(* IEC 61131-3 sources: daoli-st-library/DL_Device (part 20) *)

(* ---- FB_DL_EfEmDoorInterlockPlus.st ---- *)
(*==============================================================================
 * 组件名称 (Component)  : FB_DL_EfEmDoorInterlockPlus
 * 所属子库 (Sublibrary) : DL_Device
 * 当前版本 (Version)    : 1.0.0
 * 兼容性 (Platform)     : CODESYS 3.5 / TwinCAT 3 / 汇川 InoProShop（纯标准元素，零方言）
 * 功能描述 (Function)   : EFEM 门 / 阀 / 真空三域互斥与首因仲裁。唯一放行出口 bRelease
 *                         由四类阻断条件（门未关、阀位矛盾、真空不足、片在位）合成，阻断
 *                         域掩码逐域可见，首因只报一个编号（同拍取编号最小，锁存至复位）。
 *                         不做门体驱动输出、不做真空泵控制、不做安全回路硬线替代（安全
 *                         回路必须另有硬线双通道，本件只做逻辑侧互斥）。
 *                         门状态字位段（头注释即契约）：bit0 门关到位 ｜ bit1 门开到位 ｜
 *                         bit2 门锁到位 ｜ bit3~bit15 保留且必须为 0。
 * 溯源 (Origin)         : 道莅 clean-room 防御性实现
 * 本文件内含 (Contains) : TYPE E_DL_EfEmDomain / FUNCTION_BLOCK FB_DL_EfEmDoorInterlockPlus
 * 依赖 (Depends)        : 无（纯布尔/浮点防御逻辑，仅 Standard.library 的 ABS）
 * 红线自检 (Redline)    : 无外部全局变量、无硬件地址直引 ｜ 全变量中英双语同行注释
 *                         真空门限判零防除零 ｜ 真空非有限按保守侧（真空不足）处理 ｜
 *                         阀位矛盾判定前置于互斥仲裁 ｜ 枚举显式赋值 ｜ CASE 含 ELSE 兜底
 *                         本件无定时器/沿实例，故无周期刷新项（结构上无条件分支）
 * 错误码表 (Codes)      : 16#0003_03AC 就绪（放行或禁用，无故障）
 *                         16#0003_03AD 故障级 门状态字非法（保留位非 0）。反证句：保留位
 *                                    脏数据在输出侧与「门未关」同为禁行，不可由首因 1 区分，
 *                                    故必须独立成码
 *                         16#0003_03AE 故障级 阀位矛盾或真空门限组态非法（双反馈同 TRUE /
 *                                    同为 FALSE / 门限 ≤0）
 *                         16#0003_03AF 故障级 真空读数非有限，按「真空不足」保守侧禁行
 *                         16#0003_03B0 预留：本版不发码（下一轮区间起点，禁止回填）
 * 修订历史 (Revision)   : 2026-11-17  v1.0.0  首版入库 · R28 · 阶段三批 1
 * 验收向量 (Acceptance) : 正向 门关（状态字 bit0=1、bit2=1）、阀开反馈有效、真空 0.1 kPa
 *                         低于门限 5 kPa → 禁行、首因 3、掩码 bit2；抽到 0.05 kPa →
 *                         放行、首因清零
 *                         反向 阀双反馈同为 FALSE → 16#0003_03AE 且禁行；真空给 NaN →
 *                         16#0003_03AF 且按真空不足禁行（首因 3）；门限给 0 → 16#0003_03AE；
 *                         状态字保留位 bit7 置 1 → 16#0003_03AD 且禁行
 *============================================================================*)

(*-----------------------------------------------------------------------------
 * 枚举: E_DL_EfEmDomain（归属本功能块，同文件发布，全库唯一定义）
 * 含义: 首因所属域，每个成员在 CASE 中有且仅有一个标签。
 *----------------------------------------------------------------------------*)
TYPE E_DL_EfEmDomain :
(
    eNone    := 0,    // 无阻断域：三域全放行 / No blocking domain, all domains released
    eDoor    := 1,    // 门域：门未关到位 / Door domain, the door is not closed
    eValve   := 2,    // 阀域：阀位矛盾 / Valve domain, contradictory valve position
    eVacuum  := 3,    // 真空域：真空不足或读数非有限 / Vacuum domain, insufficient vacuum or a non-finite reading
    eWafer   := 4,    // 片域：腔内片在位（E84 语义） / Wafer domain, a wafer is present inside the chamber
    eIllegal := 99    // 非法域：状态字保留位非 0 / Illegal domain, reserved bits of the status word are set
);
END_TYPE

FUNCTION_BLOCK FB_DL_EfEmDoorInterlockPlus
VAR_INPUT
    bEnable         : BOOL := FALSE;      // 使能，FALSE 即禁行（失效导向安全侧） / Enable, FALSE forces the release output off
    uDoorStatusWord : WORD;               // 门状态字 [bit]，bit0 关到位 bit1 开到位 bit2 锁到位 bit3~15 保留 / Door status word
    bValveClosed    : BOOL := FALSE;      // 阀关到位反馈 / Valve closed feedback
    bValveOpened    : BOOL := FALSE;      // 阀开到位反馈 / Valve opened feedback
    fVacuum_kPa     : REAL := 101.3;      // 腔体真空 [kPa(abs)]，域 0~101.3 / Chamber vacuum in kilopascal absolute, domain 0 to 101.3
    fVacuumOk_kPa   : REAL := 5.0;        // 允许开门真空门限 [kPa(abs)] / Vacuum threshold permitting the door to open
    bWaferPresent   : BOOL := FALSE;      // 腔内片在位（E84 语义） / Wafer present in the chamber
    bReset          : BOOL := FALSE;      // 首因与锁存复位，上升沿生效 / First-cause and latch reset, rising edge
END_VAR
VAR_OUTPUT
    bRelease        : BOOL;               // 三域放行（唯一出口） / Three-domain release, the single outlet
    bDoorPermit     : BOOL;               // 允许开门（与放行同源，语义收窄为门域） / Door open permit, same source as the release
    uFirstCause     : UINT;               // 首因编号 1 门未关 2 阀位矛盾 3 真空不足 4 片在位 [—] / First cause number
    uBlockMask      : WORD;               // 阻断域掩码 bit0 门 bit1 阀 bit2 真空 bit3 片 [bit] / Blocking domain mask
    bError          : BOOL;               // 故障级标志，仅故障级码置位 / Fault-class flag, set on fault codes only
    eErr            : UDINT;              // 错误码，段位 16#0003_xxxx / Error code in segment 16#0003_xxxx
END_VAR
VAR
    _bInit          : BOOL := FALSE;      // 首扫标志，取非判定 / First-scan flag, tested negated
    _bDoorClosed    : BOOL;               // 门关到位（状态字 bit0） / Door closed, status word bit 0
    _bLocked        : BOOL;               // 门锁到位（状态字 bit2） / Door locked, status word bit 2
    _bReservedBad   : BOOL;               // 状态字保留位非 0 / Reserved bits of the status word are set
    _bValveBad      : BOOL;               // 阀位矛盾 / Contradictory valve position
    _bVacBad        : BOOL;               // 真空不足（含读数非有限） / Insufficient vacuum including non-finite readings
    _bCfgBad        : BOOL;               // 真空门限组态非法 / Vacuum threshold configuration invalid
    _bBlkDoor       : BOOL;               // 门域阻断 / Door domain blocked
    _bBlkValve      : BOOL;               // 阀域阻断 / Valve domain blocked
    _bBlkVac        : BOOL;               // 真空域阻断 / Vacuum domain blocked
    _bBlkWafer      : BOOL;               // 片域阻断 / Wafer domain blocked
    _bAnyBlock      : BOOL;               // 任一域阻断 / Any domain blocked
    _bFirstLatched  : BOOL;               // 首因已锁存（锁存后不再改判） / First cause latched and no longer re-arbitrated
    _eDomain        : E_DL_EfEmDomain := E_DL_EfEmDomain.eNone; // 当前首因域 / Current first-cause domain
    _rtrigReset     : R_TRIG;             // 复位上升沿 / Rising edge of the reset command
END_VAR
VAR CONSTANT
    DL_EFEM_READY      : UDINT := 16#0003_03AC;  // 就绪码 / Ready code
    DL_EFEM_WORD_BAD   : UDINT := 16#0003_03AD;  // 故障级状态字非法码 / Fault code for an illegal status word
    DL_EFEM_VALVE_BAD  : UDINT := 16#0003_03AE;  // 故障级阀位矛盾或组态非法码 / Fault code for a valve contradiction or bad configuration
    DL_EFEM_VAC_BAD    : UDINT := 16#0003_03AF;  // 故障级真空非有限码 / Fault code for a non-finite vacuum reading
    DL_EFEM_VAC_LO     : REAL := 0.0;            // 真空物理下限 [kPa(abs)] / Physical vacuum lower bound
    DL_EFEM_VAC_HI     : REAL := 101.3;          // 真空物理上限 [kPa(abs)] / Physical vacuum upper bound
    DL_EFEM_MASK_DOOR  : WORD := 16#0001;        // 门域掩码位 [bit] / Door domain mask bit
    DL_EFEM_MASK_VALVE : WORD := 16#0002;        // 阀域掩码位 [bit] / Valve domain mask bit
    DL_EFEM_MASK_VAC   : WORD := 16#0004;        // 真空域掩码位 [bit] / Vacuum domain mask bit
    DL_EFEM_MASK_WAFER : WORD := 16#0008;        // 片域掩码位 [bit] / Wafer domain mask bit
    DL_EFEM_WORD_RSV   : WORD := 16#FFF8;        // 状态字保留位掩码 [bit] / Reserved bit mask of the status word
    DL_EFEM_CAUSE_DOOR : UINT := 1;               // 首因 1 门未关 / First cause 1, the door is not closed
    DL_EFEM_CAUSE_VALVE : UINT := 2;              // 首因 2 阀位矛盾 / First cause 2, contradictory valve position
    DL_EFEM_CAUSE_VAC  : UINT := 3;               // 首因 3 真空不足 / First cause 3, insufficient vacuum
    DL_EFEM_CAUSE_WAFER : UINT := 4;              // 首因 4 片在位 / First cause 4, a wafer is present
END_VAR

// 段 1｜输出与单拍标志预置（放行类输出先清零：失效导向安全侧）
bRelease := FALSE;                                  // 放行出口先清 / Release outlet cleared first
bDoorPermit := FALSE;                               // 开门许可先清 / Door permit cleared first
uFirstCause := 0;                                   // 首因预清 / First cause pre-cleared
uBlockMask := 16#0000;                              // 掩码预清 / Mask pre-cleared
bError := FALSE;                                    // 故障标志预清 / Fault flag pre-cleared
eErr := 0;                                          // 错误码预清 / Error code pre-cleared

// 段 2｜沿检测无条件周期刷新（严禁置于分支内）
_rtrigReset(CLK := bReset);                         // 复位沿 / Reset edge

// 段 3｜首扫初始化（判据取非，R19）
IF NOT _bInit THEN
    _eDomain := E_DL_EfEmDomain.eNone;              // 首因域待机 / First-cause domain starts at none
    _bInit := TRUE;                                 // 首扫只做一次 / The first scan runs once
END_IF

// 段 4｜复位路径：清首因锁存（放行条件本身不清，条件仍在则同拍重新锁存）
IF _rtrigReset.Q THEN
    _bFirstLatched := FALSE;                        // 首因锁存解除 / First-cause latch released
    uFirstCause := 0;                               // 首因编号清 / First-cause number cleared
    _eDomain := E_DL_EfEmDomain.eNone;              // 首因域清 / First-cause domain cleared
END_IF

// 段 5｜门状态字解析（保留位脏数据先判，避免位段错位被当门未关）
_bDoorClosed := (uDoorStatusWord AND DL_EFEM_MASK_DOOR) <> 16#0000;   // bit0 关到位 / Bit 0, closed position reached
_bLocked := (uDoorStatusWord AND 16#0004) <> 16#0000;                 // bit2 锁到位 / Bit 2, locking position reached
_bReservedBad := (uDoorStatusWord AND DL_EFEM_WORD_RSV) <> 16#0000;   // 保留位非 0 / Reserved bits are set

// 段 6｜阀位矛盾闸（前置于互斥仲裁：矛盾状态下首因必须指阀域而不是门域）
_bValveBad := (bValveClosed AND bValveOpened) OR ((NOT bValveClosed) AND (NOT bValveOpened));

// 段 7｜真空组态与读数闸（门限判零防除零；读数非有限按真空不足保守侧）
_bCfgBad := (fVacuumOk_kPa <> fVacuumOk_kPa) OR ((fVacuumOk_kPa - fVacuumOk_kPa) <> (fVacuumOk_kPa - fVacuumOk_kPa))
         OR (fVacuumOk_kPa <= DL_EFEM_VAC_LO) OR (fVacuumOk_kPa > DL_EFEM_VAC_HI);
IF (fVacuum_kPa <> fVacuum_kPa) OR ((fVacuum_kPa - fVacuum_kPa) <> (fVacuum_kPa - fVacuum_kPa)) THEN
    _bVacBad := TRUE;                               // 读数非有限：按真空不足处理 / Non-finite reading treated as insufficient vacuum
    eErr := DL_EFEM_VAC_BAD;                        // 故障级：真空读数非有限 / Fault, non-finite vacuum reading
    bError := TRUE;
ELSE
    _bVacBad := (fVacuum_kPa > fVacuumOk_kPa);      // 真空值高于门限 = 真空不足 / A value above the threshold means insufficient vacuum
END_IF
IF _bCfgBad THEN
    eErr := DL_EFEM_VALVE_BAD;                      // 故障级：真空门限组态非法 / Fault, the vacuum threshold configuration is invalid
    bError := TRUE;
END_IF
IF _bReservedBad THEN
    eErr := DL_EFEM_WORD_BAD;                       // 故障级：状态字保留位非 0 / Fault, reserved bits of the status word are set
    bError := TRUE;
END_IF
IF _bValveBad THEN
    eErr := DL_EFEM_VALVE_BAD;                      // 故障级：阀位矛盾（先于互斥判定） / Fault, contradictory valve position checked before the arbitration
    bError := TRUE;
END_IF

// 段 8｜四域阻断判定（掩码逐域可见，首因只报一个）
_bBlkDoor := (NOT _bDoorClosed) OR (NOT _bLocked);  // 门域：关到位与锁到位缺一即阻断 / Door domain blocked unless closed and locked
_bBlkValve := _bValveBad OR _bCfgBad;               // 阀域：阀位矛盾或组态非法即阻断 / Valve domain blocked on a contradiction or bad configuration
_bBlkVac := _bVacBad OR _bCfgBad;                   // 真空域：真空不足或组态非法即阻断 / Vacuum domain blocked on insufficient vacuum or bad configuration
_bBlkWafer := bWaferPresent;                        // 片域：腔内片在位即阻断 / Wafer domain blocked while a wafer is present
_bAnyBlock := _bBlkDoor OR _bBlkValve OR _bBlkVac OR _bBlkWafer;   // 任一域阻断 / Any domain blocked
IF _bBlkDoor THEN
    uBlockMask := uBlockMask OR DL_EFEM_MASK_DOOR;  // 门域掩码置位 / Door domain mask bit set
END_IF
IF _bBlkValve THEN
    uBlockMask := uBlockMask OR DL_EFEM_MASK_VALVE; // 阀域掩码置位 / Valve domain mask bit set
END_IF
IF _bBlkVac THEN
    uBlockMask := uBlockMask OR DL_EFEM_MASK_VAC;   // 真空域掩码置位 / Vacuum domain mask bit set
END_IF
IF _bBlkWafer THEN
    uBlockMask := uBlockMask OR DL_EFEM_MASK_WAFER; // 片域掩码置位 / Wafer domain mask bit set
END_IF

// 段 9｜首因仲裁（仅未锁存时仲裁；顺序 1→4 即同拍取编号最小）
IF (NOT _bFirstLatched) AND _bAnyBlock THEN
    IF _bBlkDoor THEN
        _eDomain := E_DL_EfEmDomain.eDoor;          // 优先 1：门未关 / Priority 1, the door is not closed
    ELSIF _bBlkValve THEN
        _eDomain := E_DL_EfEmDomain.eValve;         // 优先 2：阀位矛盾 / Priority 2, contradictory valve position
    ELSIF _bBlkVac THEN
        _eDomain := E_DL_EfEmDomain.eVacuum;        // 优先 3：真空不足 / Priority 3, insufficient vacuum
    ELSE
        _eDomain := E_DL_EfEmDomain.eWafer;         // 优先 4：片在位 / Priority 4, a wafer is present
    END_IF
    _bFirstLatched := TRUE;                         // 首因锁存 / First cause latched
ELSIF (NOT _bAnyBlock) THEN
    _bFirstLatched := FALSE;                        // 阻断全消失：锁存解除（状态量随条件销号） / All blocks cleared, the latch is released
    _eDomain := E_DL_EfEmDomain.eNone;              // 首因域回无 / First-cause domain back to none
END_IF

// 段 10｜首因域映射（ENUM + CASE + ELSE 兜底）
CASE _eDomain OF
    E_DL_EfEmDomain.eNone:
        uFirstCause := 0;                           // 无首因 / No first cause
    E_DL_EfEmDomain.eDoor:
        uFirstCause := DL_EFEM_CAUSE_DOOR;          // 首因 1 / First cause 1
    E_DL_EfEmDomain.eValve:
        uFirstCause := DL_EFEM_CAUSE_VALVE;         // 首因 2 / First cause 2
    E_DL_EfEmDomain.eVacuum:
        uFirstCause := DL_EFEM_CAUSE_VAC;           // 首因 3 / First cause 3
    E_DL_EfEmDomain.eWafer:
        uFirstCause := DL_EFEM_CAUSE_WAFER;         // 首因 4 / First cause 4
    E_DL_EfEmDomain.eIllegal:
        uFirstCause := 0;                           // 非法域不报首因，由 03AD 表达 / The illegal domain reports no first cause, 03AD carries it
        eErr := DL_EFEM_WORD_BAD;                   // 故障级：非法域 / Fault, illegal domain
        bError := TRUE;
    ELSE
        // 非法枚举值兜底（故障级，状态字非法码承载）
        uFirstCause := 0;
        eErr := DL_EFEM_WORD_BAD;                   // 故障级：枚举越界 / Fault, the enumeration is out of range
        bError := TRUE;
        _eDomain := E_DL_EfEmDomain.eIllegal;
END_CASE

// 段 11｜放行出口（唯一出口；使能跌落即禁行，故障级存在亦禁行）
bRelease := bEnable AND (NOT _bAnyBlock) AND (NOT _bReservedBad) AND (NOT _bCfgBad) AND (NOT _bValveBad) AND (NOT _bVacBad);
bDoorPermit := bRelease;                            // 开门许可与放行同源 / Door permit shares the release source
IF bRelease THEN
    eErr := DL_EFEM_READY;                          // 就绪：三域放行 / Ready, all domains released
ELSE
    IF NOT bEnable THEN
        eErr := DL_EFEM_READY;                      // 禁用为正常停机（掩码已标全阻断域） / Disable is a normal stop, the mask shows the blocked domains
    END_IF
END_IF
END_FUNCTION_BLOCK

(* ---- FB_DL_ElectricLinearActuator.st ---- *)
(*
  ==================================================================
  组件名 Component  : FB_DL_ElectricLinearActuator
  分类   Category   : DL_Device
  复杂度 Complexity  : cx5
  版本   Version    : 1.0.0
  功能   Purpose    : 电动推杆驱动。无位置反馈，纯时间 / 电流双模到位判定：
                      限位开关反馈模（任一端限位反馈触发）与电流堵转模（电
                      流持续超堵转阈值 tStallDebounce 消抖判到位）并联，任
                      一判据先到即停并锁存到位指示；硬过流立即脱扣；全程
                      超时保护；双输出互锁绝不同得电。
  来源   Source     : t2-2-lbp（三段分层骨架）
  溯源   Origin     : IEC 61131-3 标准语义的道莅防御性实现；电动推杆堵转
                      电流判到位与限位互锁为行业公知工程语义，clean-room
                      自研实现，未复制 LBP 或任何厂商私有库源码。
  平台   Platform   : 纯 IEC 61131-3（Standard.library: TON / R_TRIG，无私有库）
  分工声明 Split     : 与 DL_Device 存量 FB_DL_DolMotor / FB_DL_SoftStarterDrive
                      分工——两者为电机启动家族（驱动器封装），本件为直线
                      执行机构（推杆本体行程与堵转管理），不做接触器 / 晶闸
                      管启动家族语义。
  作者   Author     : 道莅代码库 · PLC 编程专家（R58）
  ------------------------------------------------------------------
  边界 Boundary     :
                      一 组态域：fCurNomA > 0（非有限闸覆盖），fCurStallMul
                         > 1.0，fCurHiMul > fCurStallMul（硬过流阈值高于堵转
                         阈值，R100 配比约束），tStrokeMax > T#0S，tStallDebounce
                         ≥ T#0S（取零为电流模禁用，仅限位模）；
                      二 双模并联：限位反馈与电流堵转任一先到即到位停机，
                         到位指示锁存至反向运动或复位沿；
                      三 双命令同拍拒绝（复位优先 = 安全侧不动作，静默拒
                         绝不置故障，本拍双输出全断）；
                      四 运动相电流非有限（R151 组态域闸全覆盖）判传感失效
                         故障级；复位沿作用域：清故障锁存 / 清到位指示 / 迁
                         空闲（三项逐项声明，解除路径 = bReset 上升沿 R188）；
                      五 无全局变量、无外部变量声明、无物理地址寻址。
  修订记录 Revision  :
    2026-11-21  v1.0.0  R58 首版（批 2 · 序号 8）
  ==================================================================
*)

TYPE E_DL_ElaPhase :
(
    eElaIdle := 0,  // 空闲：消化命令，双输出断开 / idle, both outputs off
    eElaExt  := 10, // 伸出中：正转输出得电 / extending, the forward output on
    eElaRet  := 20, // 缩回中：反转输出得电 / retracting, the reverse output on
    eElaFault:= 90  // 故障锁存：双输出安全侧断开 / the latched fault, both outputs off on the safe side
);
END_TYPE

TYPE E_DL_ElaCause :
(
    eNone          := 0, // 无成因 / no cause
    eCfgBad        := 1, // 组态非法：电流标称 / 倍数配比 / 时间窗越域（故障级，与 bError 配对）/ an illegal config
    eCurBad        := 2, // 运动相电流非有限（传感失效，故障级，与 bError 配对）/ a non finite current in motion
    eCurOverHard   := 3, // 硬过流立即脱扣（故障级，与 bError 配对）/ a hard overcurrent trip
    eStrokeTimeout := 4, // 全程超时（故障级，与 bError 配对）/ a stroke timeout
    ePhaseBad      := 5  // 非法相位兜底（故障级，与 bError 配对）/ an illegal phase fallback
);
END_TYPE

FUNCTION_BLOCK FB_DL_ElectricLinearActuator
VAR_INPUT
    bCmdExt        : BOOL := FALSE;  // 伸出命令电平 [-] / the extend command level
    bCmdRet        : BOOL := FALSE;  // 缩回命令电平 [-] / the retract command level
    bLimExtFbk     : BOOL := FALSE;  // 伸出限位开关反馈，TRUE = 已达伸出端 [-] / the extend limit feedback, true = at the extend end
    bLimRetFbk     : BOOL := FALSE;  // 缩回限位开关反馈，TRUE = 已达缩回端 [-] / the retract limit feedback, true = at the retract end
    fMotCurA       : LREAL := 0.0;   // 电机电流实测 [安培] / the motor current actual [ampere]
    fCurNomA       : LREAL := 4.0;   // 标称运行电流 [安培]，域 大于 0 / the nominal running current [ampere], above zero
    fCurStallMul   : LREAL := 1.5;   // 堵转判定倍数 [倍]，域 大于 1.0 / the stall verdict multiplier, above one
    fCurHiMul      : LREAL := 2.5;   // 硬过流倍数 [倍]，域 大于堵转倍数 / the hard overcurrent multiplier, above the stall multiplier
    tStrokeMax     : TIME := T#30S;  // 全程最大时间窗 [毫秒] / the full stroke max window [millisecond]
    tStallDebounce : TIME := T#300MS; // 堵转消抖窗 [毫秒]，取零禁用电流模 / the stall debounce window, zero disables the current mode
    bEnable        : BOOL := TRUE;   // 使能，失能双输出安全侧断开并迁空闲 [-] / enable, disabling opens both outputs and returns idle
    bReset         : BOOL := FALSE;  // 复位上升沿清故障锁存 [-] / reset rising edge clears the fault latch
END_VAR
VAR_OUTPUT
    bOutExt   : BOOL := FALSE; // 电机正转输出（仅伸出相）[-] / the forward output, the extend phase only
    bOutRet   : BOOL := FALSE; // 电机反转输出（仅缩回相）[-] / the reverse output, the retract phase only
    bInPosExt : BOOL := FALSE; // 伸出到位指示（锁存至反向或复位）[-] / the extend in position latch
    bInPosRet : BOOL := FALSE; // 缩回到位指示（锁存至反向或复位）[-] / the retract in position latch
    bArrByCur : BOOL := FALSE; // 本次到位由电流堵转模判定的指示 [-] / the arrival by the current mode indicator
    ePhase    : E_DL_ElaPhase := E_DL_ElaPhase.eElaIdle; // 相位出口 [枚举] / the phase outlet
    eCause    : E_DL_ElaCause := E_DL_ElaCause.eNone; // 成因出口，锁存回放 [枚举] / the cause outlet replayed
    bError    : BOOL := FALSE; // 故障锁存标志 [-] / the fault latch flag
END_VAR
VAR
    rtReset  : R_TRIG; // 复位沿检测，段 0 无条件刷新 / the reset edge
    tonStroke: TON;    // 全程时间窗，段 0 无条件刷新 / the stroke window
    tonStall : TON;    // 堵转消抖窗，段 0 无条件刷新 / the stall debounce window
    _ePhase  : E_DL_ElaPhase := E_DL_ElaPhase.eElaIdle; // 内部相位，CASE 唯一写入目标 / the internal phase
    _eFaulC  : E_DL_ElaCause := E_DL_ElaCause.eNone; // 故障级成因，锁存至复位沿 / the fault cause latched
    _bFault  : BOOL := FALSE; // 故障锁存位 [-] / the fault latch bit
    _bCfgOk  : BOOL := FALSE; // 组态域内 [-] / the config inside the domain
    _bInit   : BOOL := FALSE; // 首扫初始化完成标志（R310）/ the first scan flag
    _lrStall : LREAL;  // 堵转电流阈值工作量 [安培] / the stall threshold work value
    _lrHi    : LREAL;  // 硬过流阈值工作量 [安培] / the hard overcurrent threshold work value
END_VAR

// 段 0｜定时器与沿检测无条件周期刷新（禁入分支，FB50-1）/ segment 0, the unconditional refresh
rtReset(CLK := bReset); // 复位沿 / the reset edge
tonStroke(IN := ((_ePhase = E_DL_ElaPhase.eElaExt) OR (_ePhase = E_DL_ElaPhase.eElaRet)) AND (NOT _bFault) AND bEnable, PT := tStrokeMax); // 全程窗，IN 串载能相闸（纯相驻留，R145）/ the stroke window on the powered phases
tonStall(IN := ((_ePhase = E_DL_ElaPhase.eElaExt) OR (_ePhase = E_DL_ElaPhase.eElaRet)) AND (NOT _bFault) AND bEnable AND (_lrStall > 0.0) AND (fMotCurA > _lrStall), PT := tStallDebounce); // 堵转消抖窗（电流模使能且超阈）/ the stall debounce window, the current mode enabled and above the threshold

// 段 1｜首扫初始化（R310）/ segment 1, the first scan
IF NOT _bInit THEN // 首扫一拍 / the first scan
    _bInit := TRUE; // 置首扫标志 / raise the flag
END_IF

// 段 2｜复位沿作用域：清故障锁存 / 清到位指示 / 迁空闲（三项逐项声明，边界四）/ segment 2, the reset edge scope
IF rtReset.Q THEN // 复位沿 / the reset edge
    _bFault := FALSE; // 作用域一：清故障锁存 / scope one, clear the fault latch
    _eFaulC := E_DL_ElaCause.eNone; // 作用域一：清成因 / scope one, clear the cause
    bInPosExt := FALSE; // 作用域二：清伸出到位 / scope two, clear the extend latch
    bInPosRet := FALSE; // 作用域二：清缩回到位 / scope two, clear the retract latch
    bArrByCur := FALSE; // 作用域二：清电流模指示 / scope two, clear the current mode flag
    _ePhase := E_DL_ElaPhase.eElaIdle; // 作用域三：迁空闲相 / scope three, back to idle
END_IF

// 段 3｜组态域闸（边界一，R151 全覆盖：电流标称非有限 + 倍数配比 + 时间窗）/ segment 3, the config gate
_bCfgOk := (fCurNomA = fCurNomA) AND ((fCurNomA - fCurNomA) = (fCurNomA - fCurNomA)) // 标称电流非有限双判据 / the nominal current finiteness
        AND (fCurNomA > 0.0) // 标称电流域 / the nominal domain
        AND (fCurStallMul > 1.0) // 堵转倍数域 / the stall multiplier domain
        AND (fCurHiMul > fCurStallMul) // 硬过流高于堵转配比（R100）/ the hard above the stall pairing
        AND (tStrokeMax > T#0S) // 全程窗域 / the stroke window domain
        AND (tStallDebounce >= T#0S); // 消抖窗域（零 = 电流模禁用）/ the debounce domain, zero disables the current mode
IF NOT _bCfgOk THEN // 组态越域 / a config violation
    IF NOT _bFault THEN // 未锁存才迁移（锁存回放 R152）/ migrate only while unlatched
        _bFault := TRUE; // 置故障锁存 / raise the fault latch
        _eFaulC := E_DL_ElaCause.eCfgBad; // 故障级成因（R45 配对）/ the fault cause
        _ePhase := E_DL_ElaPhase.eElaFault; // 迁故障相（锁存与迁相同分支，FB50-1）/ migrate to the fault phase
    END_IF
END_IF
_lrStall := fCurNomA * fCurStallMul; // 堵转阈值（组态闸已证有限正值）/ the stall threshold
_lrHi := fCurNomA * fCurHiMul; // 硬过流阈值 / the hard threshold

// 段 4｜运动相电流域闸与硬过流监视（优先级最高，R146 按方向分列）/ segment 4, the current gate and the hard overcurrent monitor
IF (_ePhase = E_DL_ElaPhase.eElaExt) OR (_ePhase = E_DL_ElaPhase.eElaRet) THEN // 载能相 / a powered phase
    IF (fMotCurA <> fMotCurA) OR ((fMotCurA - fMotCurA) <> (fMotCurA - fMotCurA)) THEN // 电流非有限（边界四）/ a non finite current
        IF NOT _bFault THEN // 未锁存才迁移 / migrate only while unlatched
            _bFault := TRUE; // 置故障锁存 / raise the fault latch
            _eFaulC := E_DL_ElaCause.eCurBad; // 故障级成因（R45 配对）/ the fault cause
            _ePhase := E_DL_ElaPhase.eElaFault; // 迁故障相 / migrate to the fault phase
        END_IF
    ELSIF (fMotCurA > _lrHi) AND (NOT _bFault) THEN // 硬过流立即脱扣（超重侧安全立即终止，R146）/ a hard overcurrent trips immediately
        _bFault := TRUE; // 置故障锁存 / raise the fault latch
        _eFaulC := E_DL_ElaCause.eCurOverHard; // 故障级成因（R45 配对）/ the fault cause
        _ePhase := E_DL_ElaPhase.eElaFault; // 迁故障相 / migrate to the fault phase
    END_IF
END_IF

// 段 5｜相位机：ENUM + CASE，含 ELSE 非法相位兜底（R128）/ segment 5, the phase machine
CASE _ePhase OF

E_DL_ElaPhase.eElaIdle: // 空闲相：评估命令（边界三双命令同拍拒绝）/ the idle phase, the command evaluation
    IF NOT bEnable THEN // 失能驻留 / dwell while disabled
        _ePhase := E_DL_ElaPhase.eElaIdle; // 停摆驻留 / dwell
    ELSIF bCmdExt AND bCmdRet THEN // 双命令同拍拒绝（复位优先）/ the dual commands rejected
        _ePhase := E_DL_ElaPhase.eElaIdle; // 静默拒绝双输出断（本拍由出口段全断）/ a silent refusal, both outputs off this scan
    ELSIF bCmdExt THEN // 伸出命令 / an extend command
        IF bLimExtFbk THEN // 已在伸出端（拒绝移动，刷新到位指示）/ already at the extend end
            bInPosExt := TRUE; // 到位指示保持 / hold the in position latch
            _ePhase := E_DL_ElaPhase.eElaIdle; // 驻留 / dwell
        ELSE // 允许伸出 / the extend allowed
            bInPosRet := FALSE; // 清反向到位 / clear the reverse latch
            bArrByCur := FALSE; // 清电流模指示 / clear the current mode flag
            _ePhase := E_DL_ElaPhase.eElaExt; // 迁伸出相 / migrate to the extend phase
        END_IF
    ELSIF bCmdRet THEN // 缩回命令 / a retract command
        IF bLimRetFbk THEN // 已在缩回端 / already at the retract end
            bInPosRet := TRUE; // 到位指示保持 / hold the in position latch
            _ePhase := E_DL_ElaPhase.eElaIdle; // 驻留 / dwell
        ELSE // 允许缩回 / the retract allowed
            bInPosExt := FALSE; // 清反向到位 / clear the extend latch
            bArrByCur := FALSE; // 清电流模指示 / clear the current mode flag
            _ePhase := E_DL_ElaPhase.eElaRet; // 迁缩回相 / migrate to the retract phase
        END_IF
    END_IF

E_DL_ElaPhase.eElaExt: // 伸出相：双模到位判定（边界二）/ the extend phase, the dual mode arrival
    IF NOT bEnable THEN // 失能即停（R191 降级显式：输出断 + 回空闲，无故障）/ a disable stops without a fault
        _ePhase := E_DL_ElaPhase.eElaIdle; // 回空闲相 / back to idle
    ELSIF bLimExtFbk THEN // 限位模到位 / the arrival by the limit mode
        bInPosExt := TRUE; // 锁存到位指示 / latch the in position
        _ePhase := E_DL_ElaPhase.eElaIdle; // 回空闲相 / back to idle
    ELSIF tonStall.Q THEN // 电流堵转模到位（消抖窗满）/ the arrival by the stall mode
        bInPosExt := TRUE; // 锁存到位指示 / latch the in position
        bArrByCur := TRUE; // 记电流模判定指示 / raise the current mode flag
        _ePhase := E_DL_ElaPhase.eElaIdle; // 回空闲相 / back to idle
    ELSIF tonStroke.Q THEN // 全程超时（故障级）/ the stroke timeout, fault grade
        _bFault := TRUE; // 置故障锁存 / raise the fault latch
        _eFaulC := E_DL_ElaCause.eStrokeTimeout; // 故障级成因（R45 配对）/ the fault cause
        _ePhase := E_DL_ElaPhase.eElaFault; // 迁故障相 / migrate to the fault phase
    END_IF

E_DL_ElaPhase.eElaRet: // 缩回相：双模到位判定（边界二）/ the retract phase, the dual mode arrival
    IF NOT bEnable THEN // 失能即停 / a disable stops without a fault
        _ePhase := E_DL_ElaPhase.eElaIdle; // 回空闲相 / back to idle
    ELSIF bLimRetFbk THEN // 限位模到位 / the arrival by the limit mode
        bInPosRet := TRUE; // 锁存到位指示 / latch the in position
        _ePhase := E_DL_ElaPhase.eElaIdle; // 回空闲相 / back to idle
    ELSIF tonStall.Q THEN // 电流堵转模到位 / the arrival by the stall mode
        bInPosRet := TRUE; // 锁存到位指示 / latch the in position
        bArrByCur := TRUE; // 记电流模判定指示 / raise the current mode flag
        _ePhase := E_DL_ElaPhase.eElaIdle; // 回空闲相 / back to idle
    ELSIF tonStroke.Q THEN // 全程超时（故障级）/ the stroke timeout, fault grade
        _bFault := TRUE; // 置故障锁存 / raise the fault latch
        _eFaulC := E_DL_ElaCause.eStrokeTimeout; // 故障级成因（R45 配对）/ the fault cause
        _ePhase := E_DL_ElaPhase.eElaFault; // 迁故障相 / migrate to the fault phase
    END_IF

E_DL_ElaPhase.eElaFault: // 故障相：成因锁存，等复位沿；双输出安全侧断开 / the fault phase
ELSE // 非法相位兜底（R128）/ the illegal phase fallback
    _bFault := TRUE; // 置故障锁存 / raise the fault latch
    _eFaulC := E_DL_ElaCause.ePhaseBad; // 故障级成因（R45 配对）/ the fault cause
    _ePhase := E_DL_ElaPhase.eElaFault; // 迁故障相 / migrate to the fault phase
END_CASE

// 段 6｜统一出口：双输出互锁 + 故障覆盖（边界二三）/ segment 6, the unified outlet with the interlock
bOutExt := (_ePhase = E_DL_ElaPhase.eElaExt) AND bEnable AND (NOT _bFault); // 正转输出仅伸出相（互锁）/ the forward output, the extend phase only
bOutRet := (_ePhase = E_DL_ElaPhase.eElaRet) AND bEnable AND (NOT _bFault); // 反转输出仅缩回相（互锁）/ the reverse output, the retract phase only
ePhase := _ePhase; // 相位出口单点映射 / the phase outlet
IF _bFault THEN // 故障锁存优先 / the fault latch first
    eCause := _eFaulC; // 成因锁存回放（R152）/ the cause replayed
ELSE // 无锁存 / no latch
    eCause := E_DL_ElaCause.eNone; // 无成因 / no cause
END_IF
bError := _bFault; // 故障标志与锁存位同源（R191 名实双出口）/ the flag shares the latch
END_FUNCTION_BLOCK

(* ---- FB_DL_ElectrodeTabBendCtrl.st ---- *)
(*
  FB_DL_ElectrodeTabBendCtrl  —  极耳折弯角度与回弹补偿 / Electrode tab bend control with springback learning
  分类 Category : DL_Device
  码位 Code     : 16#03_2_13
  段位说明      : 03_2 段低半字节 00~0F 已满（05 为历史空穴留存），进位 13 段续号（R192）
  版本 Version  : 1.0.2
  来源 Source   : t2-2-lbp — IEC 61131-3 标准语义的道莅防御性实现
  溯源 Origin   : clean-room 实现，卷对卷极耳折弯公开工艺语义，未复制任何源码行
                  （与 FB_DL_RollerGapAdjust 分工：本件按「角度—回弹」双变量收敛；间隙调整由 RollerGapAdjust 承载）
  功能 Function : 1) 单向逼近：压头只发 CmdExtend（只进不退，防反向回弹迟滞），到位后测角；
                  2) 误差超 fAngleTolDeg 则按 fLearnGain 修正回弹学习值再弯一次，累计学习值限幅 [0, fSpringbackMaxDeg]；
                  3) 下发弯折角 fCmdAngleDeg = 目标角 + 回弹学习值；迭代收敛（|测角 − 目标| <= 容差）进 Done；
                  4) fLearnGain = 0 时学习值冻结（组态可关学习）。
  边界 Boundary : ① fTargetAngleDeg <= 0 或 > fAngleMaxDeg 判组态错；容差/迭代数/限幅/超时非法同判；
                  ② iPressCyl.bFault 判气缸故障进 Fault；步超 tStepTimeout 同判（安全侧回退）；
                  ③ 迭代数超 nMaxIteration 置 bIterationExhausted 且 bInTolerance := FALSE（不静默当作 OK，判废）；
                  ④ 回弹学习值跨批次掉电不保（本件不持非易失，持久化由上层承载）；
                  ⑤ 测角由 VAR_INPUT fAngleMeasDeg 注入（上位角度传感器，规格未列的必要引脚补充）；
                  ⑥ 解除式自证：bIterationExhausted 解除 = bReset 上升沿 AND eState = Idle（引脚可满足）；
                  ⑦ CASE 全态覆盖 + ELSE 兜底置故障相。
  依赖 Depends  : I_DL_Cylinder（注入，不实例化）；语义对齐 FB_DL_RateLimiter / FB_DL_ToleranceWindow（已注册，不实例化）
  码表 Error codes（本件格 03_2_13，子码步进 +0x100）:
    16#0003_0113 信息级：弯折迭代收敛（Done 相）
    16#0003_0213 故障级：组态非法（目标角越域 / 容差 <= 0 / 增益越 0..1 / 迭代 < 1 / 限幅 <= 0 / 超时 <= 0）
    16#0003_0313 故障级：气缸故障或步超时（逼近/测量两相独立计时），锁存至复位
    16#0003_0413 故障级：迭代耗尽判废（bIterationExhausted，bInTolerance = FALSE）
    16#0003_0513 故障级：状态机落 ELSE 兜底（非法相位 ID）

R39 返修（R38 终审挂账闭环，v1.0.2）: ① tonStep 三相共享无迁移断拍 → 拆分为三相独立实例
  （tonStepAppr 逼近超时 / tonHold 保压计时 / tonStepMeas 测量超时，IN 单相等式，跨相迁移拍必断，R228-A 达标）；
  ② eBend 复用超时计时作保压 → 保压计时改由独立实例 tonHold 承载（PT 沿用 tStepTimeout 参数，
  对外接口不变约束下保持 v1.0.1 保压时长口径；测量相补步超时保护，码 0313 覆盖口径随之扩全三相）；
  ③ eFault 无迁出 → eFault 相新增 bReset 上升沿迁出边回 eIdle（迁出条件 = 输入引脚 rtReset.Q，恒可达）。
  修订历史 Revision :
    2026-11-19  v1.0.2  R39 返修：三相 TON 拆分 + 保压分实例 + eFault 迁出边（R38 挂账三项闭环）
    2026-11-18  v1.0.0  R38 首版
*)

TYPE E_DL_TabBendState :
(
    eIdle     := 0,    // 空闲：等启动指令 / Idle, waiting for start
    eApproach := 10,   // 逼近：压头伸出至弯折位 / Approach, cylinder extending
    eBend     := 20,   // 弯折：保压至测角稳定 / Bend, pressing hold
    eMeasure  := 30,   // 测量：采测角并判收敛 / Measure, sampling angle
    eCorrect  := 40,   // 修正：更新回弹学习值 / Correct, updating learned springback
    eDone     := 50,   // 完成：收敛或判废落定 / Done, converged or scrapped
    eFault    := 90    // 故障：组态/气缸/超时锁定 / Fault, latched
);
END_TYPE

FUNCTION_BLOCK FB_DL_ElectrodeTabBendCtrl
VAR_INPUT
    bStart             : BOOL := FALSE;     // 启动指令（上升沿）/ Start command
    fAngleMeasDeg      : REAL := 0.0;       // 测角输入 [deg]（上位传感器注入）/ Measured angle input
    fTargetAngleDeg    : REAL := 90.0;      // 目标弯折角 [deg]，域 (0, fAngleMaxDeg] / Target bend angle
    fSpringbackInitDeg : REAL := 0.0;       // 初始回弹量 [deg]，域 [0, fSpringbackMaxDeg] / Initial springback
    fSpringbackMaxDeg  : REAL := 10.0;      // 回弹学习值限幅 [deg]，域 > 0 / Springback learning clamp
    fAngleMaxDeg       : REAL := 135.0;     // 目标角上限 [deg]，域 > 0 / Target angle ceiling
    fAngleTolDeg       : REAL := 0.5;       // 角度容差 [deg]，域 > 0 / Angle tolerance
    fLearnGain         : REAL := 0.5;       // 学习增益 [无量纲 0..1]，0 = 冻结学习 / Learning gain, 0 freezes
    nMaxIteration      : INT  := 5;         // 最大迭代数 [次]，域 >= 1 / Max iterations
    tStepTimeout       : TIME := T#3S;      // 单步超时 [ms]，域 > 0 / Step timeout
    bReset             : BOOL := FALSE;     // 复位（判废解除路径之一）/ Reset
END_VAR
VAR_OUTPUT
    fCmdAngleDeg          : REAL;           // 下发弯折角 [deg] = 目标 + 回弹 / Commanded bend angle
    fMeasAngleDeg         : REAL;           // 测角出口 [deg] / Measured angle outlet
    fSpringbackLearnedDeg : REAL;           // 回弹学习值 [deg] / Learned springback
    bInTolerance          : BOOL;           // 收敛在容差内 / Within tolerance
    bIterationExhausted   : BOOL;           // 迭代耗尽判废锁存 / Iteration exhausted latch
    nIteration            : INT;            // 当前迭代数 [次] / Iteration count
    nErrId                : UDINT;          // 事件码，0 = 无事件 / Event code
    eState                : E_DL_TabBendState;  // 状态出口，段尾单点映射 / State outlet
END_VAR
VAR_IN_OUT
    iPressCyl : I_DL_Cylinder;              // 压装气缸引用（注入，不实例化）/ Press cylinder reference
END_VAR
VAR
    tonStepAppr: TON;                       // 逼近相超时计时（单相独占）/ Approach timeout timer
    tonHold    : TON;                       // 保压相计时（单相独占，PT=tStepTimeout 口径）/ Bend hold timer
    tonStepMeas: TON;                       // 测量相超时计时（单相独占）/ Measure timeout timer
    tonFaultWch: TON;                       // 故障观察窗，自复位 / Fault watch window, self-resetting
    rtStart    : R_TRIG;                    // 启动上升沿 / Start rising edge
    rtReset    : R_TRIG;                    // 复位上升沿 / Reset rising edge
    _eState    : E_DL_TabBendState := E_DL_TabBendState.eIdle;   // 内部相位（CASE 唯一写入目标）/ Internal phase
    _rLearn    : REAL;                      // 回弹学习值内部量 / Internal learned springback
    _rErr      : REAL;                      // 角度误差暂存 [deg] / Angle error scratch
    _uFault    : UDINT;                     // 故障码锁存 / Latched fault code
    _uInfo     : UDINT;                     // 信息码，每拍重算 / Info code
    _bFault    : BOOL;                      // 故障锁存位 / Latched fault bit
    _bCfgBad   : BOOL;                      // 组态非法聚合 / Configuration invalid aggregate
    _bExhaust  : BOOL;                     // 迭代耗尽锁存（解除式）/ Iteration exhausted latch
END_VAR
VAR CONSTANT
    DL_WatchPt : TIME := T#2S;   // 故障观察窗 [ms]，自复位 / Fault watch window
END_VAR

(* —— 段 0：定时器与边沿无条件周期刷新（R182：调用语句不得置于 IF/CASE 内） —— *)
rtStart(CLK := bStart);                                          // 启动上升沿，每拍必调
rtReset(CLK := bReset);                                          // 复位上升沿，每拍必调
tonFaultWch(IN := (NOT tonFaultWch.Q), PT := DL_WatchPt);        // 观察窗自复位（表达式入参）
tonStepAppr(IN := (_eState = E_DL_TabBendState.eApproach), PT := tStepTimeout);  // 逼近超时（单相独占）
tonHold(IN := (_eState = E_DL_TabBendState.eBend), PT := tStepTimeout);          // 保压计时（单相独占，PT=保压口径）
tonStepMeas(IN := (_eState = E_DL_TabBendState.eMeasure), PT := tStepTimeout);   // 测量超时（单相独占）

(* —— 段 1：单拍量预清零（锁存量 _uFault/_bFault/_bExhaust/_rLearn 不入清单，R187①） —— *)
_uInfo := 16#0000_0000;         // 信息码每拍重算
bInTolerance := FALSE;          // 收敛出口缺省 FALSE（Done 相单点置位）
bIterationExhausted := _bExhaust;   // 判废出口 = 解除式锁存量（禁同拍抹除）
_bCfgBad := FALSE;              // 组态非法预清零
nErrId := 16#0000_0000;         // 事件码缺省无事件

(* —— 段 2：组态域闸（覆盖全部参与判据换算的引脚，R151） —— *)
IF (fTargetAngleDeg <= 0.0) OR (fTargetAngleDeg > fAngleMaxDeg) OR (fAngleMaxDeg <= 0.0) THEN
    _bCfgBad := TRUE;           // 目标角越域
END_IF
IF (fAngleTolDeg <= 0.0) OR (fSpringbackMaxDeg <= 0.0) THEN
    _bCfgBad := TRUE;           // 容差/限幅非法
END_IF
IF (fLearnGain < 0.0) OR (fLearnGain > 1.0) THEN
    _bCfgBad := TRUE;           // 学习增益越 0..1
END_IF
IF (nMaxIteration < 1) OR (TIME_TO_DINT(tStepTimeout) <= 0) THEN
    _bCfgBad := TRUE;           // 迭代数/超时非法
END_IF
IF (fSpringbackInitDeg < 0.0) OR (fSpringbackInitDeg > fSpringbackMaxDeg) THEN
    _bCfgBad := TRUE;           // 初始回弹越域
END_IF

(* —— 段 3：复位沿（判废解除式：bReset AND eState = Idle） —— *)
IF rtReset.Q THEN
    IF _eState = E_DL_TabBendState.eIdle THEN
        _bExhaust := FALSE;     // 判废锁存清零（解除式自证路径）
        _bFault   := FALSE;     // 清故障锁存位
        _uFault   := 16#0000_0000;
        nIteration := 0;        // 迭代计数清零
    END_IF
END_IF

(* —— 段 4：下发角计算（目标 + 学习值，限幅 [0, fSpringbackMaxDeg]） —— *)
IF NOT _bCfgBad THEN
    _rLearn := MAX(0.0, MIN(_rLearn, fSpringbackMaxDeg));   // 学习值限幅（禁越界）
    fCmdAngleDeg := fTargetAngleDeg + _rLearn;              // 下发弯折角 = 目标 + 回弹
END_IF

(* —— 段 5：相位机（只做迁移与单发命令；出口在段 8） —— *)
CASE _eState OF

E_DL_TabBendState.eIdle:
    IF _bCfgBad THEN
        _uFault := 16#0003_0213;                // 故障级：组态非法
        _bFault := TRUE;                        // 锁存（复位沿可清）
        _eState := E_DL_TabBendState.eFault;
    ELSIF rtStart.Q AND (NOT _bExhaust) THEN
        _rLearn := fSpringbackInitDeg;          // 批次起步：装初始回弹量（跨批次不保持）
        nIteration := 0;                        // 迭代计数清零
        iPressCyl.CmdExtend();      // 单发伸出（单向逼近，只进不退）
        _eState := E_DL_TabBendState.eApproach; // 进逼近相
    END_IF

E_DL_TabBendState.eApproach:
    IF iPressCyl.bFault THEN
        _uFault := 16#0003_0313;                // 故障级：气缸故障
        _bFault := TRUE;
        iPressCyl.CmdStop();        // 安全侧停
        _eState := E_DL_TabBendState.eFault;
    ELSIF iPressCyl.bExtended THEN
        _eState := E_DL_TabBendState.eBend;     // 到位：进保压相
    ELSIF tonStepAppr.Q THEN
        _uFault := 16#0003_0313;                // 故障级：逼近相步超时
        _bFault := TRUE;
        iPressCyl.CmdStop();
        _eState := E_DL_TabBendState.eFault;
    END_IF

E_DL_TabBendState.eBend:
    IF iPressCyl.bFault THEN
        _uFault := 16#0003_0313;                // 故障级：气缸故障
        _bFault := TRUE;
        iPressCyl.CmdStop();
        _eState := E_DL_TabBendState.eFault;
    ELSIF tonHold.Q THEN
        _eState := E_DL_TabBendState.eMeasure;  // 保压到点：进测量相（独立实例，R228-A）
    END_IF

E_DL_TabBendState.eMeasure:
    fMeasAngleDeg := fAngleMeasDeg;             // 测角出口刷新
    _rErr := fMeasAngleDeg - fTargetAngleDeg;   // 误差 = 测角 − 目标
    IF tonStepMeas.Q THEN
        _uFault := 16#0003_0313;                // 故障级：测量相步超时（返修补全的第三相保护）
        _bFault := TRUE;
        iPressCyl.CmdStop();
        _eState := E_DL_TabBendState.eFault;
    ELSIF ABS(_rErr) <= fAngleTolDeg THEN
        bInTolerance := TRUE;                   // 收敛：容差内
        _uInfo := 16#0003_0113;                 // 信息级：迭代收敛
        iPressCyl.CmdRetract();     // 单发缩回（批次收尾）
        _eState := E_DL_TabBendState.eDone;     // 进完成相
    ELSIF nIteration >= nMaxIteration THEN
        _bExhaust := TRUE;                      // 判废锁存（不静默当作 OK）
        _uFault := 16#0003_0413;                // 故障级：迭代耗尽
        _bFault := TRUE;
        bInTolerance := FALSE;                  // 强制 FALSE（规格强制）
        iPressCyl.CmdRetract();
        _eState := E_DL_TabBendState.eDone;     // 进完成相（判废落定）
    ELSE
        _eState := E_DL_TabBendState.eCorrect;  // 未收敛未耗尽：进修正相
    END_IF

E_DL_TabBendState.eCorrect:
    IF fLearnGain > 0.0 THEN
        _rLearn := MAX(0.0, MIN(_rLearn + _rErr * fLearnGain, fSpringbackMaxDeg));   // 学习值修正并限幅
    END_IF
    nIteration := nIteration + 1;               // 迭代计数（上限守卫在 Measure 相判定）
    iPressCyl.CmdExtend();          // 单发再弯（单向逼近）
    _eState := E_DL_TabBendState.eApproach;     // 回逼近相

E_DL_TabBendState.eDone:
    IF NOT iPressCyl.bExtended THEN
        IF NOT _bExhaust THEN
            _eState := E_DL_TabBendState.eIdle;     // 缩回完成且非判废：回空闲
        ELSE
            _eState := E_DL_TabBendState.eIdle;     // 判废也回空闲（bReset 沿清判废锁存）
        END_IF
    END_IF

E_DL_TabBendState.eFault:
    IF rtReset.Q THEN                           // 迁出边：bReset 上升沿（R228-B：输入引脚，恒可达）
        _bFault := FALSE;                       // 清故障锁存位
        _uFault := 16#0000_0000;                // 清锁存码
        _bExhaust := FALSE;                     // 判废锁存清零（迁出统一清账）
        _eState := E_DL_TabBendState.eIdle;     // 迁出：回空闲（Idle 可达路径：故障迁出边）
    END_IF

ELSE
    _uFault := 16#0003_0513;                    // 故障级：非法相位 ID 兜底
    _bFault := TRUE;                            // 锁存
    _eState := E_DL_TabBendState.eFault;        // 强制回故障相

END_CASE

(* —— 段 6：出口单点映射（名实同源；锁存码回放，禁同拍抹除） —— *)
bIterationExhausted := _bExhaust;               // 判废出口 = 锁存量（置位同拍不被抹）
IF _bFault THEN
    nErrId := _uFault;              // 故障锁存码回放
    bInTolerance := FALSE;          // 故障相收敛出口强制 FALSE（安全侧）
ELSE
    nErrId := _uInfo;               // 信息码
END_IF
eState := _eState;                  // 状态出口单点映射

END_FUNCTION_BLOCK

(* ---- FB_DL_ElectrolyteMoistureGuard.st ---- *)
//==============================================================================
// 功能块：FB_DL_ElectrolyteMoistureGuard ｜ 中文名称：注液间露点/湿度联锁（首因锁定）
// 所属子库：DL_Device ｜ 版本：v1.0.0 ｜ 兼容：CODESYS V3.5+ / TwinCAT 3 / 汇川 InoProShop
// 功能描述：电解液注液间环境联锁——露点 > 露点上限 或 相对湿度 > 湿度
//           上限，任一越限持续 tDebounce → 禁止注液（bDosingPermit :=
//           FALSE），并按「首因锁定」原则记录首个触发的判据通道（bFirstCauseDp
//           / bFirstCauseRh，锁存至 bReset，中途恢复不抹除首因——归因
//           证据链不得被后续波动重写，R81 还原方向不饱和同理）。接近
//           限值预警带内给信息级提示，供提前干预。露点由 Magnus-Tetens
//           内联解算（Device 不得调用 DL_Algo，见依赖纪律）。
// 开源溯源 (Origin)：道莅原创实现（参考锂电注液间露点联锁工程惯例（电芯制程湿度管控） 分类与参数域）
// 单位表：温度[摄氏度] / 露点[摄氏度] / 相对湿度[百分数] / 预警带[开] / 时间[ms]
// 错误码表：16#0003_018C 信息级（联锁恢复放行：阻塞判据消失回放行，
//           不置 bError）/ 16#0003_018D 信息级（接近限值预警带：露点
//           落入 [上限 - 预警带, 上限]，不置 bError）/ 16#0003_0363 故障级
//           （组态非法：上限/带宽域、去抖窗 <= 0 或任一输入非有限，
//           置 bError）/ 16#0003_0364 故障级（传感器交叉校验失败：解算
//           露点 > 干球 + 1 开，物理不可能，判温湿度通道异常，安全侧
//           禁止放行，置 bError——该场景不可由 0363 的组态类判据观测，
//           属运行数据独立域）/ 16#0003_0365 故障级兜底（状态机落 ELSE，
//           置 bError）
// 状态机：E_DL_MoistGuardState（四态：eIdle=0 / ePermit=10 / eBlock=20 /
//           eFault=99），CASE 含 ELSE 兜底，ELSE 置 0365 并撤放行
// 边界行为：① 组态非法 → 故障态锁存（放行安全侧 FALSE），bReset 复位；
//           ② 湿度域外钳 1~100 照算（Magnus 对数域下限保证）；③ 越限
//           消抖未满期判据消失 → 不进阻塞（防瞬时噪声断链）；④ 首因
//           锁存只在 bReset 清除，恢复放行不抹首因（归因证据链）；
//           ⑤ 未使能放行输出 FALSE 且 bValid := FALSE；⑥ 安全侧 =
//           故障/交叉失败路径放行恒 FALSE（禁止注液为安全侧）。
// 依赖纪律：Device 不得调用 DL_Algo——Magnus-Tetens 露点解算在本件内联
//           实现，常量口径（17.62/243.12）与 FC_DL_AirDensity 族一致性
//           由本件头注释承担验证责任，改动任一侧须复核另一侧。
// 修订历史：v1.0.0 2026-11-17 首版（R24 派单 · ROADMAP P1 §693）
//==============================================================================

(*------------------------------------------------------------------------------
 * 枚举: E_DL_MoistGuardState（归属本功能块，同文件发布，全库唯一定义）
 * 含义: 环境联锁相位，每个成员在 CASE 中有且仅有一个标签。
 *-----------------------------------------------------------------------------*)
TYPE E_DL_MoistGuardState :
(
    eIdle   := 0,   // 空闲：未使能 / Idle, not enabled
    ePermit := 10,  // 放行：判据全部满足 / Permit, all criteria satisfied
    eBlock  := 20,  // 阻塞：越限去抖确认，禁止注液 / Block, violation debounced, dosing forbidden
    eFault  := 99   // 故障：组态非法/交叉校验/非法状态 / Fault, config, cross-check or illegal state
);
END_TYPE

FUNCTION_BLOCK FB_DL_ElectrolyteMoistureGuard
VAR_INPUT
    bEnable      : BOOL;                    // 联锁使能 [—] / Interlock enable
    bReset       : BOOL;                    // 故障复位 [—]，上升沿清首因/组态锁存 / Fault reset, rising edge clears latches
    bDosingReq   : BOOL;                    // 注液请求 [—]（联锁仅门控，不接管请求） / Dosing request, gated only
    fRoomTempC   : LREAL;                   // 注液间干球温度 [摄氏度] / Room dry-bulb temperature [degC]
    fRhPct       : LREAL;                   // 注液间相对湿度 [百分数]，域外钳 1..100 照算 / Room relative humidity [percent], clamped 1..100
    fDpLimitC    : LREAL := -40.0;          // 露点联锁上限 [摄氏度]，高于此越限 / Dew-point interlock limit [degC]
    fRhLimitPct  : LREAL := 10.0;           // 湿度联锁上限 [百分数]，高于此越限，按工艺卡组态 / Humidity interlock limit [percent]
    fWarnBandK   : LREAL := 2.0;            // 接近限值预警带宽 [开]，须 >= 0 / Warning band width [K]
    tDebounce    : TIME  := T#5S;           // 越限去抖窗 [ms]，须 > 0 / Violation debounce window [ms]
END_VAR
VAR_OUTPUT
    bDosingPermit  : BOOL;                  // 注液放行 [—]（联锁门控输出） / Dosing permit, gated output
    fDewPointC     : LREAL;                 // 解算露点 [摄氏度]（诊断出口） / Solved dew point [degC], diagnostics outlet
    bFirstCauseDp  : BOOL;                  // 首因锁存：露点通道 [—]（bReset 才清除） / First-cause latch, dew-point channel
    bFirstCauseRh  : BOOL;                  // 首因锁存：湿度通道 [—]（bReset 才清除） / First-cause latch, humidity channel
    eGuardState    : E_DL_MoistGuardState;  // 联锁相位 [—] / Interlock phase
    eErr           : UDINT;                 // 错误码，0 = 无错，码位 16#0003_018C 起信息级、16#0003_0363 起故障级（分带见错误码表） / Error code, 0 = no error, band info/fault per the code table
    bError         : BOOL;                  // 故障级标志，仅故障级错误置位 / Fault-class flag, set only on fault-level codes
    bValid         : BOOL;                  // 输出可用标志 / Outputs usable flag
END_VAR
VAR
    fbDebounce : TON;                       // 越限去抖计时（每拍无条件刷新）[ms] / Violation debounce timer, refreshed unconditionally
    _eState    : E_DL_MoistGuardState := E_DL_MoistGuardState.eIdle; // 当前相位 / Current phase
    _bCfgBad   : BOOL;                      // 组态非法锁存 / Illegal config latch
    _bCrossBad : BOOL;                      // 交叉校验失败锁存 / Cross-check fault latch
    _bInfoRel  : BOOL;                      // 恢复放行信息当拍标志 / Recovery info flag of this scan
    _bInfoWarn : BOOL;                      // 预警带信息当拍标志 / Warning-band info flag of this scan
    _fRhUse    : LREAL;                     // 生效湿度（已钳位）[百分数] / Effective humidity, clamped
    _fGamma    : LREAL;                     // 露点解算中间量 ln(RH/100) [无量纲] / Dew-point intermediate
    _fDpCalc   : LREAL;                     // 解算露点 [摄氏度] / Solved dew point [degC]
    _bViolate  : BOOL;                      // 越限电平（去抖窗条件） / Violation level, debounce condition
    _bIllegal  : BOOL;                      // 非法状态标志 / Illegal state flag
    _bInit     : BOOL := FALSE;             // 首扫标志，初值 FALSE 取非判定 / First-scan flag, tested negated
END_VAR
VAR CONSTANT
    DL_EMG_MAGNUS_A : LREAL := 17.62;       // Magnus 系数 A [无量纲]，与 FC_DL_AirDensity 同口径 / Magnus coefficient A, aligned
    DL_EMG_MAGNUS_B : LREAL := 243.12;      // Magnus 系数 B [摄氏度]，同口径 / Magnus coefficient B, aligned
    DL_EMG_INF      : LREAL := 1.7976931348623157E308; // LREAL 幅值上限 / LREAL magnitude ceiling
    DL_EMG_EPS      : LREAL := 1.0E-6;      // 浮点判零容差 [混合] / Float zero tolerance
    DL_EMG_RH_MIN   : LREAL := 1.0;         // 湿度钳位下限 [百分数] / Humidity clamp floor [percent]
    DL_EMG_RH_MAX   : LREAL := 100.0;       // 湿度钳位上限 [百分数] / Humidity clamp ceiling [percent]
    DL_EMG_CROSS_K  : LREAL := 1.0;         // 交叉校验容差 [开] / Cross-check tolerance [K]
    DL_EMG_ZERO     : LREAL := 0.0;         // 零值常量，避免裸字面量 [混合] / Zero constant, avoids a bare literal
END_VAR

(*------------------------------------------------------------------------------
 * 段 1｜每拍预置：放行先断（安全侧），单拍标志预清零
 *      Permit cleared first, fail-safe, one-shot flags pre-cleared
 *-----------------------------------------------------------------------------*)
bDosingPermit := FALSE;                  // 放行先断（安全侧） / Permit cleared first
fDewPointC    := DL_EMG_ZERO;            // 露点出口先清 / Dew point cleared first
eErr   := 16#0000_0000;                  // 错误码每拍重算 / Error code recomputed
bError := FALSE;                         // 故障标志每拍重算 / Fault flag recomputed
bValid := FALSE;                         // 可用标志每拍重算 / Usable flag recomputed
_bInfoRel  := FALSE;                     // 恢复信息预清零 / Recovery info pre-cleared
_bInfoWarn := FALSE;                     // 预警信息预清零 / Warn info pre-cleared
_bIllegal  := FALSE;                     // 非法状态预清零 / Illegal flag pre-cleared

(*------------------------------------------------------------------------------
 * 段 2｜首扫初始化
 *      First-scan initialisation
 *-----------------------------------------------------------------------------*)
IF NOT _bInit THEN
    _eState    := E_DL_MoistGuardState.eIdle; // 相位空闲起步 / Phase starts idle
    _bCfgBad   := FALSE;                 // 组态锁存清零 / Config latch cleared
    _bCrossBad := FALSE;                 // 交叉锁存清零 / Cross latch cleared
    _bInit     := TRUE;                  // 首扫只做一次 / The first scan runs once
END_IF

(*------------------------------------------------------------------------------
 * 段 3｜组态防御闸：非有限（R79）+ 上限/带宽/去抖窗域
 *      Configuration defense gates
 *-----------------------------------------------------------------------------*)
IF (fRoomTempC <> fRoomTempC) OR (ABS(fRoomTempC) > DL_EMG_INF)
   OR (fRhPct <> fRhPct) OR (ABS(fRhPct) > DL_EMG_INF)
   OR (fDpLimitC <> fDpLimitC) OR (ABS(fDpLimitC) > DL_EMG_INF)
   OR (fRhLimitPct <> fRhLimitPct) OR (ABS(fRhLimitPct) > DL_EMG_INF)
   OR (fWarnBandK <> fWarnBandK) OR (ABS(fWarnBandK) > DL_EMG_INF) THEN
    _bCfgBad := TRUE;                    // 非有限归组态非法锁存 / Non-finite folded into the config latch
END_IF
IF (NOT _bCfgBad) AND ((fRhLimitPct <= DL_EMG_EPS) OR (fRhLimitPct > 100.0)
   OR (fWarnBandK < DL_EMG_ZERO) OR (tDebounce <= T#0MS)) THEN
    _bCfgBad := TRUE;                    // 上限/带宽/去抖窗域非法锁存 / Limit, band and window domains latched
END_IF
IF bReset THEN
    _bCfgBad   := FALSE;                 // 复位清组态锁存 / Reset clears the config latch
    _bCrossBad := FALSE;                 // 复位清交叉锁存 / Reset clears the cross latch
    bFirstCauseDp := FALSE;              // 复位清首因锁存（露点） / Reset clears the dew-point first cause
    bFirstCauseRh := FALSE;              // 复位清首因锁存（湿度） / Reset clears the humidity first cause
END_IF

(*------------------------------------------------------------------------------
 * 段 4｜湿度钳位与露点内联解算（Device 泳道零外部依赖）
 *      Humidity clamp and the inline dew-point solve
 *-----------------------------------------------------------------------------*)
_fRhUse := MIN(MAX(fRhPct, DL_EMG_RH_MIN), DL_EMG_RH_MAX); // 湿度双侧钳位 / Two-sided humidity clamp
_fGamma := LN(_fRhUse / 100.0);          // 中间量 ln(RH/100) [无量纲]，恒 <= 0 / Intermediate, always <= 0
_fDpCalc := DL_EMG_MAGNUS_B * _fGamma / (DL_EMG_MAGNUS_A - _fGamma); // Magnus 露点反解 [摄氏度]，分母恒 > 17 / Magnus dew-point solve
fDewPointC := _fDpCalc;                  // 露点诊断出口 / Dew-point diagnostics outlet

(*------------------------------------------------------------------------------
 * 段 5｜传感器交叉校验：露点 > 干球 + 容差 → 物理不可能，安全侧禁止放行
 *      Sensor cross-check, safe side blocks the permit
 *-----------------------------------------------------------------------------*)
IF (NOT _bCfgBad) AND (_fDpCalc > (fRoomTempC + DL_EMG_CROSS_K)) THEN
    _bCrossBad := TRUE;                  // 交叉校验失败锁存 / Cross-check failure latched
END_IF

(*------------------------------------------------------------------------------
 * 段 6｜越限电平与去抖计时无条件刷新（R40：CASE 之外每拍必调）
 *      Violation level and debounce timer refreshed unconditionally
 *-----------------------------------------------------------------------------*)
_bViolate := (_fDpCalc > fDpLimitC) OR (_fRhUse > fRhLimitPct); // 双判据任一越限 / Either criterion violated
fbDebounce(IN := (_eState = E_DL_MoistGuardState.ePermit) AND _bViolate,
           PT := tDebounce);             // 越限去抖窗（放行态起算） / Violation debounce window, from the permit phase

(*------------------------------------------------------------------------------
 * 段 7｜相位机（CASE 含 ELSE 兜底；状态改写只出现在分支判据内，R39）
 *      Phase machine with ELSE fallback
 *-----------------------------------------------------------------------------*)
IF (NOT bEnable) OR _bCfgBad OR _bCrossBad THEN
    _eState := E_DL_MoistGuardState.eFault; // 未使能或异常转故障态（放行 FALSE） / Not enabled or anomaly, fault, permit FALSE
ELSE
CASE _eState OF

    E_DL_MoistGuardState.eIdle:            // 空闲：使能进放行态
        IF bEnable THEN
            _eState := E_DL_MoistGuardState.ePermit; // 进放行 / To permit
        END_IF

    E_DL_MoistGuardState.ePermit:          // 放行：越限去抖满进阻塞；预警带提示
        IF NOT bEnable THEN
            _eState := E_DL_MoistGuardState.eFault; // 使能撤销转故障 / Enable dropped, fault
        ELSIF fbDebounce.Q THEN
            IF _fDpCalc > fDpLimitC THEN
                bFirstCauseDp := TRUE;     // 首因锁定：露点通道（bReset 才清） / First cause, dew-point channel
            END_IF
            IF _fRhUse > fRhLimitPct THEN
                bFirstCauseRh := TRUE;     // 首因锁定：湿度通道（bReset 才清） / First cause, humidity channel
            END_IF
            _eState := E_DL_MoistGuardState.eBlock; // 进阻塞 / To block
        ELSIF _fDpCalc >= (fDpLimitC - fWarnBandK) THEN
            _bInfoWarn := TRUE;            // 接近限值预警带（信息级） / Warning-band notice, info
        END_IF

    E_DL_MoistGuardState.eBlock:           // 阻塞：越限判据全部消失回放行（首因保持）
        IF NOT bEnable THEN
            _eState := E_DL_MoistGuardState.eFault; // 使能撤销转故障 / Enable dropped, fault
        ELSIF (NOT _bViolate) AND (NOT fbDebounce.Q) THEN
            _bInfoRel := TRUE;             // 联锁恢复放行（信息级，拍 N 进入） / Recovery, permit restored, info
            _eState := E_DL_MoistGuardState.ePermit; // 回放行 / Back to permit
        END_IF

    E_DL_MoistGuardState.eFault:           // 故障：复位沿且原因消失回空闲
        IF bReset AND (NOT _bCfgBad) AND (NOT _bCrossBad) THEN
            _eState := E_DL_MoistGuardState.eIdle; // 回空闲 / Back to idle
        END_IF

    ELSE                                   // 非法状态兜底（R21：CASE 必带 ELSE）
        _bIllegal := TRUE;                 // 标记非法状态 / Flag the illegal state
        _eState   := E_DL_MoistGuardState.eFault; // 回故障态（放行 FALSE） / Back to fault, permit FALSE
END_CASE
END_IF

(*------------------------------------------------------------------------------
 * 段 8｜码位出口与放行（故障级码 3 行内置 bError，R45/R101 配对）
 *      Code outlet and release, fault codes paired with bError
 *-----------------------------------------------------------------------------*)
IF _bIllegal THEN
    eErr   := 16#0003_0365;                // 故障级：状态机兜底 / Fault: state machine fallback
    bError := TRUE;                        // 置故障标志 / Raise the fault flag
ELSIF _bCrossBad THEN
    eErr   := 16#0003_0364;                // 故障级：传感器交叉校验失败 / Fault: sensor cross-check failed
    bError := TRUE;                        // 置故障标志 / Raise the fault flag
ELSIF _bCfgBad THEN
    eErr   := 16#0003_0363;                // 故障级：组态非法 / Fault: illegal configuration
    bError := TRUE;                        // 置故障标志 / Raise the fault flag
ELSIF _bInfoWarn THEN
    eErr := 16#0003_018D;                  // 信息级：接近限值预警带 / Info: warning band
ELSIF _bInfoRel THEN
    eErr := 16#0003_018C;                  // 信息级：联锁恢复放行 / Info: interlock recovery
END_IF

bDosingPermit := (NOT bError) AND (_eState = E_DL_MoistGuardState.ePermit); // 放行挂状态量（R99） / Permit bound to the state
bValid := (NOT bError) AND bEnable AND (_eState <> E_DL_MoistGuardState.eIdle); // 空闲/故障/未使能输出不可用 / Outputs unusable in idle, fault or disabled
eGuardState := _eState;                  // 相位出口 / Phase outlet
END_FUNCTION_BLOCK

(* ---- FB_DL_ElectrolyteTankLevel.st ---- *)
(*==============================================================================
 * 组件名称 (Component)  : FB_DL_ElectrolyteTankLevel
 * 溯源说明 (Provenance) : 道莅 clean-room 防御性实现（路线图 L350 已登记 + Building 族借形）
 * 所属子库 (Sublibrary) : DL_Device / TankControl
 * 当前版本 (Version)    : 1.0.0
 * 兼容性   (Platform)   : CODESYS 3.5 / TwinCAT 3 / 汇川 InoProShop；
 *                         纯 IEC 61131-3（第 3 版），零标准库依赖
 * 组件分类 (Category)   : 功能块（FUNCTION_BLOCK）· 电解液储罐液位双限 + 氮封监视
 * 功能一句话 (Summary)  : 液位双限告警 + 氮封微正压联锁 + 加注许可仲裁，仅监视与许可。
 * 边界与安全 (Boundary) : ①传感器失效 → 保持上次有效状态 + 压力故障 + 禁加注（安全侧）；
 *                         ②LoLo 大于等于 HiHi → 设定值非法码且禁加注；
 *                         ③液位高于 HiHi 禁加注，低于 LoLo 同禁（双侧禁注）；
 *                         ④氮封压力低于下限开氮阀，高于上限置越限码；
 *                         ⑤NaN 液位/压力拒收并按传感器失效处理（安全侧）。
 * 错误码    : 16#0003_037B 液位/压力传感器失效——故障级（持续态）
 *             16#0003_037C 氮封压力越限（高于上限或低于下限）——故障级（持续态）
 *             16#0003_037D 双限设定值非法（LoLo 不小于 HiHi）——故障级（持续态）
 * 码位总账  : 16#0003_037B 用 / 16#0003_037C 用 / 16#0003_037D 用
 * 修改记录  : v1.0.0 R26 初版
 *==============================================================================*)
FUNCTION_BLOCK FB_DL_ElectrolyteTankLevel
VAR_INPUT
    fLevel    : LREAL; // 液位 [%] / Level [%]
    fN2Press  : LREAL; // 氮封压力 [kPa] / Nitrogen blanket pressure [kPa]
    fHiHi     : LREAL; // 液位高高限 [%] / Level high-high limit [%]
    fLoLo     : LREAL; // 液位低低限 [%] / Level low-low limit [%]
    fPressLo  : LREAL; // 氮封压力下限 [kPa] / Pressure lower limit [kPa]
    fPressHi  : LREAL; // 氮封压力上限 [kPa] / Pressure upper limit [kPa]
    bSensorOk : BOOL;  // 传感器通道自诊断 OK / Sensor channel self-check OK
END_VAR
VAR_OUTPUT
    bFillPermit  : BOOL; // 加注许可仲裁输出 / Fill permit arbitration
    bN2ValveOpen : BOOL; // 氮封阀开建议（TRUE=建议开启）/ N2 valve open request
    bHiHi        : BOOL; // 液位高高告警 / Level high-high alarm
    bLoLo        : BOOL; // 液位低低告警 / Level low-low alarm
    bPressFault  : BOOL; // 氮封压力故障 / Nitrogen pressure fault
    eErr         : UDINT; // 本周期错误码，0=无错 / Error code this cycle, 0 = none
END_VAR
VAR
    bLevelHiHiL : BOOL; // 液位高高内部判定 / Internal high-high predicate
    bLevelLoLoL : BOOL; // 液位低低内部判定 / Internal low-low predicate
    fLevelGuard : LREAL; // 液位实时守卫副本 / Level guard copy
    fPressGuard : LREAL; // 压力实时守卫副本 / Pressure guard copy
    bParamOk    : BOOL;  // 设定值合法性 / Setpoint legality
END_VAR

// ---------- 实时守卫副本（内部判定统一用，输出为锁存结论） ----------
fLevelGuard := fLevel;
fPressGuard := fN2Press;

// ---------- 设定值防御：LoLo 不小于 HiHi 即非法（含 NaN 拒收） ----------
bParamOk := (fLoLo < fHiHi) AND (fPressLo < fPressHi)
        AND (fLoLo = fLoLo) AND (fHiHi = fHiHi) AND (fPressLo = fPressLo) AND (fPressHi = fPressHi);
IF NOT bParamOk THEN
    bFillPermit := FALSE;                     // 设定非法禁加注（安全侧）/ Illegal setpoints, no fill
    eErr := 16#0003_037D;                     // 设定非法码 / Illegal setpoints code
    RETURN;
END_IF

// ---------- 传感器防御：通道失效或 NaN 均按失效处理 ----------
IF (NOT bSensorOk) OR (fLevelGuard <> fLevelGuard) OR (fPressGuard <> fPressGuard) THEN
    // 保持上次有效状态：bHiHi/bLoLo/bN2ValveOpen 锁存值不动，禁加注与压力故障置位
    bFillPermit := FALSE;                     // 禁加注（安全侧）/ Fill forbidden, safe side
    bPressFault := TRUE;                      // 压力故障置位 / Pressure fault set
    eErr := 16#0003_037B;                     // 传感器失效码 / Sensor failure code
    RETURN;
END_IF

// ---------- 双限判定（实时值判据，输出为持续态结论） ----------
bLevelHiHiL := fLevelGuard >= fHiHi;          // 高高判据 / High-high predicate
bLevelLoLoL := fLevelGuard <= fLoLo;          // 低低判据 / Low-low predicate
bHiHi := bLevelHiHiL;                         // 对外告警（持续态）/ Alarm output
bLoLo := bLevelLoLoL;

// ---------- 氮封压力监视：低于下限开氮阀，高于上限越限 ----------
bPressFault := (fPressGuard > fPressHi) OR (fPressGuard < fPressLo); // 越限判据 / Out-of-band predicate
IF fPressGuard < fPressLo THEN
    bN2ValveOpen := TRUE;                     // 压力不足开氮阀 / Low pressure: open N2 valve
    eErr := 16#0003_037C;                     // 越限码 / Out-of-band code
ELSIF fPressGuard > fPressHi THEN
    bN2ValveOpen := FALSE;                    // 超压关氮阀 / Over pressure: close N2 valve
    eErr := 16#0003_037C;                     // 越限码（复用同码）/ Out-of-band code shared
ELSE
    bN2ValveOpen := FALSE;                    // 带内保持关闭 / In-band stays closed
END_IF

// ---------- 加注许可仲裁：双限内 + 压力正常才放行 ----------
IF bHiHi OR bLoLo OR bPressFault THEN
    bFillPermit := FALSE;                     // 任一异常禁加注 / Any anomaly forbids fill
ELSE
    bFillPermit := TRUE;                      // 全部正常放行 / All normal permits fill
END_IF

END_FUNCTION_BLOCK

(* ---- FB_DL_ElMutingGantry.st ---- *)
(*
  FB_DL_ElMutingGantry  —  EL 检测龙门进出光幕屏蔽（muting）/ EL gantry light-curtain muting arbitration
  分类 Category : DL_Device
  码位 Code     : 16#03_2_19
  段位说明      : 03_2 段低半字节已满，1x 段续号，18 格由 DoorInterlockHvac 启用，本件启用 19 格（R192）
  版本 Version  : 1.0.0
  来源 Source   : t1-5-tcopen — EL 检测龙门屏蔽时序仲裁待挖项
  溯源 Origin   : clean-room 实现，2+2 传感器 muting 为公开标准时序语义，未复制任何源码行
  功能 Function : 1) 四传感器（进向 S1/S2，出向 S3/S4）2+2 时序判进/出方向：
                  进向对 S1 先 S2 后激活 → 进向屏蔽；出向对 S3 先 S4 后激活 → 出向屏蔽；
                  2) 屏蔽窗超时 tonMuteIn/tonMuteOut 强制退出屏蔽并锁故障（防遮蔽卡死常屏蔽）；
                  3) 安全事件不受屏蔽约束之外的部分：光幕触发位仅在无屏蔽时升级为安全停止；
                  屏蔽有效期间光幕触发按正常穿越处理（标准 muting 语义）；
                  4) bMuteLamp 屏蔽指示灯出口（标准 muting 联锁灯）。
  边界 Boundary : ① 本件只做屏蔽时序仲裁，光幕本体语义由 FB_DL_SafetyLightCurtain 承载
                  （本件仅接收其触发位，不实例化、不替代）；
                  ② 双向对同时激活判组态矛盾（故障级锁存）；
                  ③ R228-A 达标声明：tonMuteIn/tonMuteOut 各自单相独占（IN 为单相等式），跨相迁移拍 IN 必断；
                  ④ R228-B 达标声明：eFault 迁出 = rtReset.Q AND NOT 双向矛盾 AND NOT 超时残留，
                  三条件均为可满足输入（矛盾解除、复位给沿后），无恒假子式，逐字写于此；
                  ⑤ 传感器经 4 只 FB_DL_SignalDebounce 消抖（主体首部无条件刷新）。
  依赖 Depends  : FB_DL_SignalDebounce（实例化 ×4）；FB_DL_SafetyLightCurtain（语义对齐，不实例化）
  码表 Error codes（本件格 03_2_19，子码步进 +0x100）:
    16#0003_0119 信息级：屏蔽窗正常退出（穿越完成）
    16#0003_0219 故障级：屏蔽窗超时强制退出（防遮蔽卡死），锁存至复位
    16#0003_0319 故障级：双向对同拍激活（组态/传感器矛盾），锁存至复位
    16#0003_0419 故障级：状态机落 ELSE 兜底（非法相位 ID），锁存至复位
    16#0003_0519 信息级：光幕触发且无屏蔽（安全停止有效，本件只透传不仲裁）

  修订历史 Revision :
    2026-11-19  v1.0.0  R39 首版（批次 3 · 序号 11）
*)

TYPE E_DL_ElMuteState :
(
    eIdle    := 0,    // 无屏蔽：等传感器时序 / Idle, no muting active
    eMuteIn  := 10,   // 进向屏蔽：S1→S2 时序命中 / Entry muting, S1 then S2 sequence
    eMuteOut := 20,   // 出向屏蔽：S3→S4 时序命中 / Exit muting, S3 then S4 sequence
    eFault   := 90    // 故障：超时/矛盾锁定 / Fault, latched
);
END_TYPE

FUNCTION_BLOCK FB_DL_ElMutingGantry
VAR_INPUT
    bS1       : BOOL := FALSE;        // 进向传感器 1（外沿）/ Entry sensor 1, outer
    bS2       : BOOL := FALSE;        // 进向传感器 2（内沿）/ Entry sensor 2, inner
    bS3       : BOOL := FALSE;        // 出向传感器 1（内沿）/ Exit sensor 1, inner
    bS4       : BOOL := FALSE;        // 出向传感器 2（外沿）/ Exit sensor 2, outer
    bCurtainTrip : BOOL := FALSE;     // 光幕触发位（FB_DL_SafetyLightCurtain 输出透传）/ Light curtain tripped passthrough
    tDebounce : TIME := T#10MS;       // 传感器消抖延时 [ms] / Sensor debounce delay
    tMuteMax  : TIME := T#10S;        // 屏蔽窗上限 [ms]，域 > 0 / Maximum muting window
    bReset    : BOOL := FALSE;        // 故障复位，上升沿生效 / Fault reset, rising edge
END_VAR
VAR_OUTPUT
    eMuteDir    : E_DL_ElMuteState;   // 屏蔽方向出口（Idle = 无屏蔽）/ Muting direction outlet
    bMuteActive : BOOL;               // 屏蔽生效中（进向或出向）[-] / Muting active flag
    bMuteLamp   : BOOL;               // 屏蔽指示灯出口（与 bMuteActive 同源）[-] / Muting lamp output
    bSafetyStop : BOOL;               // 安全停止出口：光幕触发且无屏蔽（电平，每拍重算）[-] / Safety stop output
    bError      : BOOL;               // 故障锁存，仅故障级码置位，bReset 清除 [-] / Fault latch
    uErrorId    : UDINT;              // 事件码，0 = 无事件（故障级锁存回放）/ Event code
END_VAR
VAR
    afbDeb     : ARRAY[0..3] OF FB_DL_SignalDebounce;   // 四传感器消抖实例，主体首部无条件刷新 / Sensor debounce instances
    tonMuteIn  : TON;                 // 进向屏蔽窗计时（单相独占，R228-A）/ Entry mute window timer, single phase
    tonMuteOut : TON;                 // 出向屏蔽窗计时（单相独占，R228-A）/ Exit mute window timer, single phase
    rtReset    : R_TRIG;              // 复位上升沿 / Reset rising edge
    rtS1       : R_TRIG;              // 进向 S1 上升沿（时序判向基准）/ S1 rising edge, sequence basis
    rtS3       : R_TRIG;              // 出向 S3 上升沿（时序判向基准）/ S3 rising edge, sequence basis
    i0         : INT;                 // 消抖阵列遍历索引 [0..3] / Debounce array loop index
    _eState    : E_DL_ElMuteState := E_DL_ElMuteState.eIdle;  // 内部相位（CASE 唯一写入目标）/ Internal phase
    _bS1St     : BOOL;                // S1 消抖稳定镜像 / S1 debounced mirror
    _bS2St     : BOOL;                // S2 消抖稳定镜像 / S2 debounced mirror
    _bS3St     : BOOL;                // S3 消抖稳定镜像 / S3 debounced mirror
    _bS4St     : BOOL;                // S4 消抖稳定镜像 / S4 debounced mirror
    _bSeqIn    : BOOL;                // 进向时序命中记忆（S1 沿后 S2 激活）/ Entry sequence memory
    _bSeqOut   : BOOL;                // 出向时序命中记忆（S3 沿后 S4 激活）/ Exit sequence memory
    _bFault    : BOOL;                // 故障锁存位 / Latched fault bit
    _uFault    : UDINT;               // 故障码锁存寄存 / Latched fault code register
    _uInfo     : UDINT;               // 信息码，每拍重算 / Info code
    _bConflict : BOOL;                // 双向矛盾聚合 / Bidirectional conflict aggregate
END_VAR

(* —— 段 0：定时器与边沿实例无条件周期刷新（R182：调用语句不得置于 IF/CASE 内） —— *)
FOR i0 := 0 TO 3 DO                                          // 消抖阵列每拍全量刷新（等效无条件域）
    afbDeb[i0](bRawInput := bS1 AND (i0 = 0)                 // 位选：0=S1 1=S2 2=S3 3=S4
                            OR (bS2 AND (i0 = 1))
                            OR (bS3 AND (i0 = 2))
                            OR (bS4 AND (i0 = 3)),
               tRiseDelay := tDebounce,                      // 消抖延时（组态透传）
               tFallDelay := tDebounce,
               bEnable := TRUE);
END_FOR
rtS1(CLK := afbDeb[0].bStable);                              // S1 沿（消抖后取沿）
rtS3(CLK := afbDeb[2].bStable);                              // S3 沿（消抖后取沿）
rtReset(CLK := bReset);                                      // 复位沿刷新，每拍必调
tonMuteIn(IN := (_eState = E_DL_ElMuteState.eMuteIn), PT := tMuteMax);    // 进向屏蔽窗（单相独占）
tonMuteOut(IN := (_eState = E_DL_ElMuteState.eMuteOut), PT := tMuteMax);  // 出向屏蔽窗（单相独占）

(* —— 段 1：单拍量预清零（锁存量 _uFault/_bFault/_bSeqIn/_bSeqOut 不入清单，R187①） —— *)
_uInfo := 16#0000_0000;             // 信息码每拍重算
_bConflict := FALSE;                // 双向矛盾预清零（段 3 单点聚合）
uErrorId := 16#0000_0000;           // 事件码缺省无事件

(* —— 段 2：消抖镜像采集 —— *)
_bS1St := afbDeb[0].bStable;        // S1 稳定值
_bS2St := afbDeb[1].bStable;        // S2 稳定值
_bS3St := afbDeb[2].bStable;        // S3 稳定值
_bS4St := afbDeb[3].bStable;        // S4 稳定值

(* —— 段 3：双向矛盾与故障聚合 —— *)
IF _bS1St AND _bS2St AND _bS3St AND _bS4St THEN
    _bConflict := TRUE;             // 四传感器全亮：双向矛盾（组态/遮蔽异常）
END_IF
IF _bConflict AND (NOT _bFault) THEN
    _uFault := 16#0003_0319;        // 故障级：双向同拍激活
    _bFault := TRUE;
END_IF

(* —— 段 4：时序判向记忆（进向：S1 沿先行，S2 激活命中；出向同构） —— *)
IF rtS1.Q THEN
    _bSeqIn := TRUE;                // S1 沿：进向时序开窗（由 S2 激活或对释放关闭）
END_IF
IF _bS2St AND _bSeqIn THEN
    ;                               // S2 激活且时序开窗：进向屏蔽请求在相位机判定
ELSIF (NOT _bS1St) AND (NOT _bS2St) THEN
    _bSeqIn := FALSE;               // 进向对全释放：时序记忆关闭
END_IF
IF rtS3.Q THEN
    _bSeqOut := TRUE;               // S3 沿：出向时序开窗
END_IF
IF (NOT _bS3St) AND (NOT _bS4St) THEN
    _bSeqOut := FALSE;              // 出向对全释放：时序记忆关闭
END_IF

(* —— 段 5：相位机（屏蔽仲裁；出口在段 7） —— *)
CASE _eState OF

E_DL_ElMuteState.eIdle:
    IF _bFault THEN
        _eState := E_DL_ElMuteState.eFault;         // 聚合故障直接进故障相
    ELSIF _bS1St AND _bS2St AND _bSeqIn THEN
        _eState := E_DL_ElMuteState.eMuteIn;        // 进向时序命中：进屏蔽相
    ELSIF _bS3St AND _bS4St AND _bSeqOut THEN
        _eState := E_DL_ElMuteState.eMuteOut;       // 出向时序命中：进屏蔽相
    END_IF

E_DL_ElMuteState.eMuteIn:
    IF _bFault THEN
        _eState := E_DL_ElMuteState.eFault;         // 聚合故障直接进故障相
    ELSIF tonMuteIn.Q THEN
        _uFault := 16#0003_0219;                    // 故障级：屏蔽窗超时强制退出
        _bFault := TRUE;
        _bSeqIn := FALSE;                           // 强制退出：时序记忆作废
        _eState := E_DL_ElMuteState.eFault;
    ELSIF (NOT _bS1St) AND (NOT _bS2St) THEN
        _uInfo := 16#0003_0119;                     // 信息级：进向穿越完成正常退出
        _bSeqIn := FALSE;                           // 时序记忆关闭
        _eState := E_DL_ElMuteState.eIdle;          // 回无屏蔽相
    END_IF

E_DL_ElMuteState.eMuteOut:
    IF _bFault THEN
        _eState := E_DL_ElMuteState.eFault;         // 聚合故障直接进故障相
    ELSIF tonMuteOut.Q THEN
        _uFault := 16#0003_0219;                    // 故障级：屏蔽窗超时强制退出
        _bFault := TRUE;
        _bSeqOut := FALSE;                          // 强制退出：时序记忆作废
        _eState := E_DL_ElMuteState.eFault;
    ELSIF (NOT _bS3St) AND (NOT _bS4St) THEN
        _uInfo := 16#0003_0119;                     // 信息级：出向穿越完成正常退出
        _bSeqOut := FALSE;                          // 时序记忆关闭
        _eState := E_DL_ElMuteState.eIdle;          // 回无屏蔽相
    END_IF

E_DL_ElMuteState.eFault:
    ;                               // 故障相：等复位沿（段 6 承载迁出）

ELSE
    _uFault := 16#0003_0419;        // 故障级：非法相位 ID 兜底
    _bFault := TRUE;
    _eState := E_DL_ElMuteState.eFault;             // 强制回故障相

END_CASE

(* —— 段 6：eFault 迁出沿（R228-B：rtReset.Q AND NOT 矛盾 AND NOT 超时残留，逐字自证见头注释④） —— *)
IF rtReset.Q AND (NOT _bConflict) THEN
    _bFault := FALSE;               // 清故障锁存位
    _uFault := 16#0000_0000;
    IF _eState = E_DL_ElMuteState.eFault THEN
        _eState := E_DL_ElMuteState.eIdle;          // 故障相迁出：回无屏蔽相
    END_IF
END_IF

(* —— 段 7：出口单点映射（名实同源；锁存码回放，禁同拍抹除） —— *)
bMuteActive := (_eState = E_DL_ElMuteState.eMuteIn) OR (_eState = E_DL_ElMuteState.eMuteOut);   // 屏蔽生效中
bMuteLamp := bMuteActive;           // 指示灯同源镜像
bSafetyStop := bCurtainTrip AND (NOT bMuteActive);   // 安全停止：光幕触发且无屏蔽（电平每拍重算）
IF bSafetyStop THEN
    _uInfo := 16#0003_0519;         // 信息级：安全停止有效（覆盖正常退出码，安全信息优先）
END_IF
IF _bFault THEN
    uErrorId := _uFault;            // 故障锁存码回放
    bError := TRUE;
ELSE
    uErrorId := _uInfo;             // 信息码
    bError := FALSE;
END_IF
eMuteDir := _eState;                // 方向出口单点映射

END_FUNCTION_BLOCK

(* ---- FB_DL_EmergencyStopChainDiag.st ---- *)
//==============================================================================
// 功能块：FB_DL_EmergencyStopChainDiag ｜ 中文名称：急停回路多节点诊断聚合与断链定位
// 所属子库：DL_Device ｜ 版本：v1.0.0 ｜ 日期：2026-11-23
// 兼容：CODESYS V3.5+ / TwinCAT 3 / 汇川 InoProShop（纯 IEC 61131-3 第 3 版，零方言）
// 功能描述：急停安全回路四节点（急停按钮 NC 反馈 / 双通道继电器反馈 / 回路
//           复位反馈）诊断聚合：四节点全好 → 回路完好；任一节点断 → 经去抖
//           确认后锁存断链故障并按优先级定位首个断点（按钮 > K1 > K2 > 复位），
//           复位沿且四节点恢复才解除锁存；复位沿而回路未恢复判复位时序非法
//           （信息级）。安全声明：本件只做诊断聚合与逻辑级 bSafeOut，物理
//           输出侧必须在 PRG_IoMapping 层做双保险切断（安全最高优先级拦截），
//           本件输出不得单独驱动任何安全执行器。
// 开源溯源 (Origin)：原创实现（t2-8-isa182 报警与回路诊断语义深化，零外部
//           源码行，clean-room 独立编写）
// 公开接口清单：输入 bBtnOk / bK1FbOk / bK2FbOk / bResetOk / bReset / tDebounce；
//               输出 bChainOk / bSafeOut / eBreakNode / uErrCode / bError / bValid
// 单位表：全部 BOOL / TIME 引脚，无量纲；tDebounce[ms]
// 输入契约：四节点反馈为 NC 回路完好电平（TRUE = 完好），引脚经 IO 映射层
//           注入；bReset 为操作员复位按钮沿。
// 输出契约：bSafeOut 为逻辑级安全输出（物理双保险在输出映射层）；
//           eBreakNode 锁存回放至解锁沿；uErrCode 故障级锁存、信息级每拍
//           重算；bError 仅断链故障相保持。
// 错误码表：16#0003_0760 故障级（急停回路断链，置 bError，锁存至复位沿回放）/
//           16#0003_0761 信息级（复位时序非法：复位沿而回路未恢复，不置
//           bError）/
//           16#0003_0762 预留禁用（不得挪用）
// 状态机：E_DL_EStopDiagState（本文件唯一定义，全库唯一属主）：
//           eHealthy = 0 / eBroken = 1；非法状态兜底归 eBroken（安全侧）
// 边界行为：① 断链经 tDebounce 去抖确认才锁存（反馈抖动不误报）；
//           ② 断点定位在确认瞬间按按钮→K1→K2→复位优先级单拍锁存，
//             故障期内锁存回放，不按当下输入重推断（R189）；
//           ③ 解锁条件 = 复位上升沿 AND 四节点全恢复（可达清除沿已声明）；
//           ④ TON/R_TRIG 每拍无条件刷新（不入分支，红线 R7）；
//           ⑤ 输入非有限不适用（BOOL 引脚无浮点域，域闸由组态域承担）；
//           ⑥ CASE 带 ELSE 非法态兜底归 eBroken（安全侧）。
// 修订历史：v1.0.0 2026-11-23 首版（R73 派单 · 批 1 · 序 4）
//==============================================================================

(*------------------------------------------------------------------------------
 * 枚举 1: E_DL_EStopDiagState（归属本功能块，同文件发布，全库唯一属主）
 * 含义: 诊断状态机相位，成员与 CASE 标签双向完备。
 *-----------------------------------------------------------------------------*)
TYPE E_DL_EStopDiagState :
(
    eHealthy := 0,   // 回路完好：四节点全恢复且锁存已解除 / Chain healthy, all nodes restored
    eBroken  := 1    // 断链锁存：故障码与断点回放中 / Broken, fault code and break node replaying
);
END_TYPE

(*------------------------------------------------------------------------------
 * 枚举 2: E_DL_EStopNode（归属本功能块，同文件发布，全库唯一属主）
 * 含义: 断链定位节点，eNone = 无断点。
 *-----------------------------------------------------------------------------*)
TYPE E_DL_EStopNode :
(
    eNone  := 0,   // 无断点 / No break point
    eBtn   := 1,   // 急停按钮节点断 / E-stop button node broken
    eK1    := 2,   // 安全继电器 K1 反馈节点断 / Safety relay K1 feedback node broken
    eK2    := 3,   // 安全继电器 K2 反馈节点断 / Safety relay K2 feedback node broken
    eReset := 4    // 回路复位反馈节点断 / Chain reset feedback node broken
);
END_TYPE

(*==============================================================================
 * 功能块: FB_DL_EmergencyStopChainDiag
 * 调用约定: 每个扫描周期无条件调用一次；实例状态全部驻留于私有变量。
 * 调用示例: eStopDiag(bBtnOk := NOT bEStopRawNc, bK1FbOk := bK1Mon,
 *                     bK2FbOk := bK2Mon, bResetOk := bResetLoopMon,
 *                     bReset := bAckBtn, tDebounce := T#50MS);
 *          断链定位读 eStopDiag.eBreakNode 送上位机诊断画面；bSafeOut 参与
 *          输出映射层双保险合取。
 * 组装说明: ① 安全组装纪律：物理切断通道必须由 PRG_IoMapping 层对本件
 *             bSafeOut 与硬件安全回路触点做双保险串联，本件输出单独不得
 *             驱动任何安全执行器（安全最高优先级拦截声明）；
 *           ② 四节点反馈引脚全部经 PRG_IoMapping 读入，本件零 %I/%Q
 *             物理地址（红线 R2）；
 *           ③ 复位按钮沿在本件内去抖无效——操作员复位须经 bResetOk
 *             反馈恢复后才可达解锁沿，双条件合取由 eBroken 相承担；
 *           ④ 本件可与任意数量下游工艺联锁件组合，bChainOk 作公共使能
 *             因子注入各工艺件的 bEn 合取项。
 *==============================================================================*)
FUNCTION_BLOCK FB_DL_EmergencyStopChainDiag
VAR_INPUT
    bBtnOk    : BOOL := FALSE;       // 急停按钮 NC 反馈（TRUE = 未按下/完好）/ E-stop button NC feedback, TRUE = intact
    bK1FbOk   : BOOL := FALSE;       // 安全继电器 K1 反馈（TRUE = 吸合正常）/ Safety relay K1 feedback, TRUE = healthy
    bK2FbOk   : BOOL := FALSE;       // 安全继电器 K2 反馈（TRUE = 吸合正常）/ Safety relay K2 feedback, TRUE = healthy
    bResetOk  : BOOL := TRUE;        // 回路复位反馈（TRUE = 复位回路完好）/ Reset loop feedback, TRUE = healthy
    bReset    : BOOL := FALSE;       // 操作员复位按钮（上升沿有效）/ Operator reset pushbutton, rising edge active
    tDebounce : TIME := T#50MS;      // 断链去抖确认延时 [ms] / Break debounce delay [ms]
END_VAR
VAR_OUTPUT
    bChainOk  : BOOL;                // 回路完好声明（去抖后）/ Chain healthy declaration after debounce
    bSafeOut  : BOOL;                // 逻辑级安全输出（物理双保险在 IO 映射层）/ Logic-level safe output, physical double cut at the IO mapping layer
    eBreakNode: E_DL_EStopNode;      // 断点定位（锁存回放）/ Break node location, latched replay
    uErrCode  : UDINT;               // 错误码，0 = 无错 / Error code, 0 = no error
    bError    : BOOL;                // 故障级标志，仅故障级错误置位 / Fault-class flag, set only on fault-level codes
    bValid    : BOOL;                // 输出可用标志 / Outputs usable flag
END_VAR
VAR
    tonBrk    : TON;                 // 断链去抖定时器，每拍无条件刷新 / Break debounce timer, refreshed every scan
    trigReset : R_TRIG;              // 复位沿检测，每拍无条件刷新 / Reset edge detector, refreshed every scan
    bChainRaw : BOOL;                // 四节点原始合取（未去抖）/ Raw four-node AND, not debounced
    bSeqBad   : BOOL;                // 复位时序非法声明 / Reset sequence violation flag
    eState    : E_DL_EStopDiagState; // 诊断状态机相位（私有驻留）/ Diagnostic state machine phase, private resident
END_VAR
VAR CONSTANT
    DL_ES_CODE_BRK : UDINT := 16#0003_0760; // 故障级：断链码 / Fault code: chain broken
    DL_ES_CODE_SEQ : UDINT := 16#0003_0761; // 信息级：复位时序非法码 / Info code: illegal reset sequence
END_VAR

// ---- 段 1｜定时/沿实例无条件刷新（红线 R7：禁入条件分支）----
bChainRaw := bBtnOk AND bK1FbOk AND bK2FbOk AND bResetOk; // 四节点原始合取 / Raw four-node AND
tonBrk(IN := NOT bChainRaw, PT := tDebounce);            // 断链去抖按断态断输入 / Break timer input per raw break state
trigReset(CLK := bReset);                                 // 复位沿每拍刷新 / Reset edge refreshed every scan

// ---- 段 2｜出口默认值：入口即赋确定值 ----
bChainOk := FALSE;                    // 回路完好默认 FALSE / Chain healthy preset FALSE
bSafeOut := FALSE;                    // 安全输出默认 FALSE（安全侧）/ Safe output preset FALSE, safe side
bSeqBad  := FALSE;                    // 时序非法声明先清零 / Sequence violation preset FALSE
uErrCode := 16#0000_0000;             // 信息码每拍重算（信息级不锁存，R189）/ Info code recomputed, never latched per R189
bError   := FALSE;                    // 故障标志先清零（故障相由锁存改写）/ Fault flag cleared, overwritten by latch in the fault phase
bValid   := TRUE;                     // 可用标志默认 TRUE / Usable flag preset TRUE

// ---- 段 3｜诊断状态机（CASE 带 ELSE；断点锁存单拍定位）----
CASE eState OF
    E_DL_EStopDiagState.eHealthy:     // 完好相：监视断链
        bChainOk := TRUE;             // 完好声明 / Healthy declared
        bSafeOut := bChainRaw;        // 安全输出随原始合取（去抖前透传，断后去抖确认才翻）/ Safe out follows raw AND
        IF tonBrk.Q THEN              // 断链去抖确认（可达进入沿）/ Break confirmed by debounce
            eState := E_DL_EStopDiagState.eBroken; // 进入断链锁存相 / Enter the broken latch phase
            IF NOT bBtnOk THEN        // 断点定位：按钮优先 / Locate: button first
                eBreakNode := E_DL_EStopNode.eBtn;
            ELSIF NOT bK1FbOk THEN    // 次优先 K1 / Then K1
                eBreakNode := E_DL_EStopNode.eK1;
            ELSIF NOT bK2FbOk THEN    // 次优先 K2 / Then K2
                eBreakNode := E_DL_EStopNode.eK2;
            ELSE                      // 余下为复位反馈节点 / Remaining: reset feedback node
                eBreakNode := E_DL_EStopNode.eReset;
            END_IF
            uErrCode := DL_ES_CODE_BRK; // 故障码锁存（回放至解锁）/ Fault code latched, replayed until release
            bError   := TRUE;           // 置故障标志（R45 配对）/ Raise the fault flag, R45 pairing
        ELSIF trigReset.Q THEN        // 完好态复位沿为无效时序 / Reset edge while healthy is a sequence violation
            bSeqBad  := TRUE;         // 信息级留痕 / Info-level trace
            uErrCode := DL_ES_CODE_SEQ; // 信息级：复位时序非法（不置 bError）/ Info: illegal reset sequence, no fault flag
        END_IF

    E_DL_EStopDiagState.eBroken:      // 断链锁存相：故障码与断点回放
        bChainOk := FALSE;            // 回路不完好声明 / Chain unhealthy declared
        bSafeOut := FALSE;            // 安全输出切断（安全侧）/ Safe output cut, safe side
        bError   := TRUE;             // 故障级锁存回放 / Fault-class latch replay
        uErrCode := DL_ES_CODE_BRK;   // 故障码回放（不在故障相重推断）/ Fault code replayed, never re-inferred
        IF trigReset.Q THEN           // 复位沿处理（锁存声明的清除沿）/ Reset edge, the declared release edge
            IF bChainRaw THEN         // 四节点全恢复才允许解锁 / All nodes restored before release
                eState := E_DL_EStopDiagState.eHealthy; // 回完好相 / Back to the healthy phase
                eBreakNode := E_DL_EStopNode.eNone;     // 断点定位清零 / Break node cleared
                uErrCode   := 16#0000_0000;             // 故障码清零 / Fault code cleared
                bError     := FALSE;                    // 故障标志解除 / Fault flag released
            ELSE
                bSeqBad  := TRUE;     // 回路未恢复时的复位判时序非法 / Reset while broken is a sequence violation
                uErrCode := DL_ES_CODE_SEQ; // 信息级留痕（故障码保持回放）/ Info trace, fault code keeps replaying
                bError   := TRUE;     // 故障级保持 / Fault class held
            END_IF
        END_IF

    ELSE                              // 非法状态兜底（R21：CASE 必带 ELSE）
        eState   := E_DL_EStopDiagState.eBroken; // 拦截非法值归断链（安全侧）/ Catch illegal value to broken, safe side
        bSafeOut := FALSE;            // 安全输出切断 / Safe output cut
        bError   := TRUE;             // 兜底相按故障级处理 / Fallback phase treated as fault class
        uErrCode := DL_ES_CODE_BRK;   // 兜底故障码 / Fallback fault code
END_CASE

bValid := TRUE;                       // 全部出口确定：输出可用 / All outlets deterministic, outputs usable
END_FUNCTION_BLOCK
